(* IEC 61131-3 sources: daoli-st-library/DL_Process (part 2) *)

(* ---- FB_DL_ColumnDpCtrl.st ---- *)
(*==============================================================================
 * 组件名称 (Component)  : FB_DL_ColumnDpCtrl
 * 溯源说明 (Provenance): 道莅 clean-room 防御性实现（IEC 61131-3 纯净实现，闭源文档仅借语义，零代码行）
 * 所属子库 (Sublibrary) : DL_Process / ProcessControl
 * 当前版本 (Version)    : 1.0.0
 * 兼容性   (Platform)   : CODESYS 3.5 / TwinCAT 3 / 汇川 InoProShop / 施耐德
 *                         Machine Expert；纯 IEC 61131-3（第 3 版），仅用
 *                         Standard.library 的 TON / LIMIT / ABS / TIME_TO_DINT / DINT_TO_TIME
 * 组件分类 (Category)   : 功能块（FUNCTION_BLOCK）· 精馏塔压差控制
 * 功能一句话 (Summary)  : 以塔压差设定为基准增量式双向调节回流与再沸两路给定，
 *                         带死区、双侧抗饱和，压差越上限时按防冲塔策略强制分配。
 *
 * 本件存在的意义 (Why this unit exists)
 *   精馏塔的 ΔP 是「液泛前兆」的直接指示：ΔP 升高说明上升蒸汽被液相托住，
 *   继续加热会冲塔（产品全部跑废、可能超压）。库内 FB_DL_RatioController 管
 *   两路比值、FB_DL_SplitRangeControl 管单输出分程，都不解「ΔP 偏高时增回流
 *   减再沸、ΔP 偏低时反向」这条双向分配律，也没有防冲塔的强制优先级。
 *
 * 增量式调节与抗饱和 (Incremental law and anti-windup)
 *   两路输出都是**增量累加**的绝对给定（不是增量输出），每走一步：
 *     ΔP 偏高（> 设定 + 死区）→ 回流 +fStep、再沸 −fStep
 *     ΔP 偏低（< 设定 − 死区）→ 回流 −fStep、再沸 +fStep
 *   累加后钳到 fOutMin~fOutMax，且**到达限值即停止向该方向累加**——钳位后
 *   不再累加是本件的抗饱和手段，不做积分回算（塔的工艺时间常数以十分钟计，
 *   回算没有收益，只会让审计算不清）。
 *
 * 防冲塔优先级 (Anti-flooding priority)
 *   fDpMeas > fDpHighLimit 持续 tConfirm → bDpHigh：**再沸立即降到 fOutMin、
 *   回流抬到 fOutMax**，压差调节暂时让位。这条优先级高于增量调节，因为冲塔
 *   是不可逆的产品损失；退出须压差回落到 fDpHighLimit − fDpDeadband 以下
 *   （用已有死区引脚做回差，不新开参数），避免在限值上反复进出。
 *
 * 引脚补全声明 (Pin completion —— 规格正文要求但引脚表漏列)
 *   fStep : 单步调节量 [%]，规格正文明确要求「步长引脚 fStep（缺省 1.0 %）」；
 *   tStep : 步进节拍 [ms]，增量式调节必须有时基，否则步进率随任务周期漂移。
 *   tStep 采用 T#200MS 缺省（现场常规回路周期），两引脚均已按要求常量化默认值。
 *
 * 边界安全 (Boundary)
 *   ① fDpSp <= 0、fOutMin >= fOutMax、fDpHighLimit <= fDpSp、fStep <= 0、
 *      任一参数非有限 → 故障 030E、**双输出置 fOutMin**（切断热源侧再加量）；
 *   ② fDpMeas 非有限 → 故障 030F、**保持末次输出**（塔不能因坏值断热，
 *      与①方向相反，两条并列写死）；
 *   ③ 死区内 → 信息 01DC，不调节、输出保持；
 *   ④ bDpHigh 进入置 01DD，退出复用 01DC（R90 不加码，头注释写明复用理由）；
 *   ⑤ 失能 → eIdle、双输出置 fOutMin、bDpHigh 清零（逐项赋，R72）；
 *   ⑥ 两只 TON 无条件刷新（步进节拍 / 越限确认），各司其职不共用；
 *   ⑦ CASE 落 ELSE 置 0310 并回 eFault。
 *
 * 错误码    : 16#0005_01DC ΔP 在死区内不调节，或已退出防冲塔——信息级，正常调节
 *             16#0005_01DD ΔP 越上限，已按防冲塔策略强制分配——信息级，保护动作
 *             16#0005_030E 控制参数非法（设定/限值/步长/上下限关系）——故障级，双输出置下限
 *             16#0005_030F ΔP 输入非有限，保持末次输出——故障级，不得断热
 *             16#0005_0310 状态机落 ELSE 兜底（非法状态）——故障级，回 eFault
 * 码位总账  : 16#0005_01DC 用 / 16#0005_01DD 用 ｜ 16#0005_030E 用 / 16#0005_030F 用 / 16#0005_0310 用
 * 状态机    : E_DL_ColumnDpState（eIdle / eNormal / eDpHigh / eDpLow / eFault），CASE 含 ELSE 兜底，
 *             ELSE 置 16#0005_0310 并回 eFault；失能无条件回 eIdle
 * 采样约定  : 每任务周期调用一次；步进节拍由 tStep 给定，越限确认由 tConfirm 给定
 * 依赖说明  : 只做组合编排，不复制低层算法；无 DL_ 子库调用
 * 验收向量  : V1 ΔP 5.0、设定 5.0、死区 0.2 → 死区内不调节，eErr = 01DC，输出保持
 *             V2 ΔP 6.0（> 5.2）、步长 1.0、节拍 200 ms → 每步回流 +1、再沸 −1，
 *                累加到限值后停（抗饱和主向量）
 *             V3 V2 持续到回流 = fOutMax → bLimited = TRUE，不再向该方向累加
 *             V4 ΔP 8.5（> 上限 8.0）持续 2 s → bDpHigh = TRUE，回流 = fOutMax、
 *                再沸 = fOutMin，eErr = 01DD（防冲塔主向量）
 *             V5 V4 后 ΔP 回落到 7.9（< 8.0 − 0.2）→ 退出防冲塔，eErr = 01DC（回差主向量）
 *             V6 fDpSp = 0 → 030E，双输出 = fOutMin，bValid = FALSE
 *             V7 fDpMeas = NaN → 030F，双输出保持上一拍值（坏值不断热主向量）
 *             V8 bEnable 落 → eIdle，双输出 = fOutMin，bDpHigh = FALSE
 * 红线自检  : 全局变量声明零使用 / 外部变量访问零使用 / 物理地址零使用 ｜ 纯 IEC 61131-3 ｜ 无除法
 *             浮点只用大小与容差比较 ｜ 无循环 ｜ 全变量双语同行注释 ｜ ENUM + CASE
 *             含 ELSE ｜ 两只 TON 在主体前部无条件刷新 ｜ 阈值常量化，无魔法数
 * 修订历史  : 2026-11-16  v1.0.0  首版入库（R22 · 批 3 · 过程单元控制）
 *============================================================================*)

(*-----------------------------------------------------------------------------
 * 枚举: E_DL_ColumnDpState（归属本功能块，同文件发布，全库唯一定义）
 * 含义: 塔压差控制相位。0 起步长 10。
 *-----------------------------------------------------------------------------*)
TYPE E_DL_ColumnDpState :
(
    eIdle   := 0,      // 待机：未使能或参数非法 / Idle, disabled or illegal parameters
    eNormal := 10,     // 正常：ΔP 在死区外按增量调节 / Normal, incremental control outside the dead band
    eDpHigh := 20,     // 压差高：防冲塔强制分配 / High differential pressure, anti-flooding distribution
    eDpLow  := 30,     // 压差低：反向调节 / Low differential pressure, reverse correction
    eFault  := 99      // 故障：参数非法或输入非有限 / Fault, illegal parameter or non-finite input
);
END_TYPE

FUNCTION_BLOCK FB_DL_ColumnDpCtrl
VAR_INPUT
    fDpMeas      : REAL;                       // 塔压差实测 [kPa] / measured column differential pressure [kPa]
    fDpSp        : REAL := 5.0;                // 压差设定 [kPa]，须 > 0 / differential pressure setpoint [kPa], must be > 0
    fDpDeadband  : REAL := 0.2;                // 死区半宽 [kPa]，须 >= 0 / dead band half width [kPa], must be >= 0
    fOutMin      : REAL := 0.0;                // 输出下限 [%] / output floor [%]
    fOutMax      : REAL := 100.0;              // 输出上限 [%]，须 > fOutMin / output ceiling [%], must exceed the floor
    fDpHighLimit : REAL := 8.0;                // 防冲塔压差上限 [kPa]，须 > fDpSp / anti-flooding limit [kPa], must exceed the setpoint
    fStep        : REAL := 1.0;                // 单步调节量 [%]，须 > 0 / single step size [%], must be > 0
    tStep        : TIME := T#200MS;            // 步进节拍 [ms] / step cadence [ms]
    tConfirm     : TIME := T#2S;               // 越限确认时间 [ms] / limit confirm time [ms]
    bEnable      : BOOL;                       // 使能 / enable
END_VAR
VAR_OUTPUT
    fRefluxOut   : REAL;                       // 回流量给定 [%]，范围 fOutMin~fOutMax / reflux setpoint [%]
    fReboilOut   : REAL;                       // 再沸热源给定 [%]，范围 fOutMin~fOutMax / reboiler duty setpoint [%]
    bDpHigh      : BOOL;                       // 压差越上限（防冲塔生效） / differential pressure above the limit
    bLimited     : BOOL;                       // 输出已到限值（抗饱和生效） / an output sits at its limit
    eErr         : UDINT;                      // 错误码，0 表示无错 / error code, 0 means no error
    bError       : BOOL;                       // 故障级标志，仅故障级错误置位 / fault-class flag, set only on fault-level codes
    bValid       : BOOL;                       // 输出可用标志 / outputs usable flag
END_VAR
VAR
    fbStep       : TON;                        // 步进节拍计时，段 6 无条件刷新 [ms] / step cadence timer
    fbHigh       : TON;                        // 越限确认计时，段 6 无条件刷新 [ms] / limit confirm timer
    _eState      : E_DL_ColumnDpState := E_DL_ColumnDpState.eIdle; // 当前相位 / current phase
    _bInit       : BOOL := FALSE;              // 首扫标志，初值 FALSE 取非判定 / first-scan flag, tested negated
    _bParamBad   : BOOL;                       // 参数非法标志 / illegal parameter flag
    _bFiniteBad  : BOOL;                       // 输入非有限标志 / non-finite input flag
    _bIllegal    : BOOL;                       // 非法状态标志 / illegal state flag
    _bStepBreak  : BOOL;                       // 步进计时器断输入一拍 / step timer one-scan break
    _bHighBreak  : BOOL;                       // 越限计时器断输入一拍 / limit timer one-scan break
    _bStepPulse  : BOOL;                       // 本拍走一步 / one step this scan
    _bInDeadband : BOOL;                       // 本拍在死区内 / inside the dead band this scan
    _bHiAbove    : BOOL;                       // 本拍越上限（裸判据） / above the limit this scan
    _bHiExit     : BOOL;                       // 压差已回落到退出线以下 / below the exit line
    _tStepUse    : TIME := T#200MS;            // 生效步进节拍 [ms]，已钳位 / effective cadence, clamped
    _tConfUse    : TIME := T#2S;               // 生效确认时间 [ms]，已钳位 / effective confirm time, clamped
    _fReflux     : REAL;                       // 回流量累加保持量 [%] / held reflux setpoint [%]
    _fReboil     : REAL;                       // 再沸累加保持量 [%] / held reboiler setpoint [%]
    _fRefluxOut  : REAL;                       // 回流输出暂存 [%] / reflux outlet staging
    _fReboilOut  : REAL;                       // 再沸输出暂存 [%] / reboiler outlet staging
END_VAR
VAR CONSTANT
    DL_VAL_LIM     : REAL := 1.0E6;            // 有限性判定的绝对值上限 [无量纲] / finiteness ceiling
    DL_SP_MIN      : REAL := 0.0;              // 设定下限 [kPa]，须严格大于 / setpoint floor, strictly greater
    DL_BAND_MIN    : REAL := 0.0;              // 死区下限 [kPa] / dead band floor [kPa]
    DL_STEP_MIN    : REAL := 0.0;              // 步长下限 [%]，须严格大于 / step floor, strictly greater
    DL_EPS         : REAL := 1.0E-6;           // 浮点比较容差 [%] / float comparison tolerance [%]
    DL_CAD_MIN_MS  : DINT := 10;               // 步进节拍下限 [ms] / cadence floor [ms]
    DL_CAD_MAX_MS  : DINT := 60000;            // 步进节拍上限 [ms] / cadence ceiling [ms]
    DL_CONF_MAX_MS : DINT := 60000;            // 确认时间上限 [ms] / confirm ceiling [ms]
    DL_TIME_ZERO   : TIME := T#0MS;            // 时间零值基准 [ms] / time zero reference
END_VAR

(*------------------------------------------------------------------------------
 * 段 1｜每拍预置（输出与累加量在段 9 单点写入）
 *      Per-scan presets, the outputs and accumulators are written in segment nine
 *-----------------------------------------------------------------------------*)
eErr         := 16#0000_0000;                  // 错误码每拍重算 / error code recomputed every scan
bError       := FALSE;                         // 故障标志每拍重算 / fault flag recomputed every scan
bValid       := FALSE;                         // 可用标志每拍重算 / usable flag recomputed every scan
bDpHigh      := FALSE;                         // 越限标志每拍重算 / high flag recomputed
bLimited     := FALSE;                         // 抗饱和标志每拍重算 / limited flag recomputed
_bParamBad   := FALSE;                         // 参数非法标志预清零 / parameter flag pre-cleared
_bFiniteBad  := FALSE;                         // 非有限标志预清零 / non-finite flag pre-cleared
_bIllegal    := FALSE;                         // 非法状态标志预清零 / illegal state flag pre-cleared
_bStepPulse  := FALSE;                         // 步进脉冲预置 FALSE / step pulse preset FALSE
_bInDeadband := FALSE;                         // 死区标志预置 FALSE / dead band flag preset FALSE
_bHiAbove    := FALSE;                         // 越上限标志预置 FALSE / above-limit preset FALSE
_bHiExit     := FALSE;                         // 退出标志预置 FALSE / exit preset FALSE

(*------------------------------------------------------------------------------
 * 段 2｜首扫初始化（两路从输出下限起：塔未运行时回流与热源都在最小位）
 *      First-scan initialisation, both loops start at the output floor
 *-----------------------------------------------------------------------------*)
IF NOT _bInit THEN
    _eState     := E_DL_ColumnDpState.eIdle;   // 相位待机 / phase idle
    _fReflux    := 0.0;                        // 回流累加量 0 [%] / reflux accumulator zero
    _fReboil    := 0.0;                        // 再沸累加量 0 [%] / reboiler accumulator zero
    _bStepBreak := TRUE;                       // 步进节拍从零开始 / cadence timer starts from zero
    _bHighBreak := TRUE;                       // 越限确认从零开始 / confirm timer starts from zero
    _bInit      := TRUE;                       // 首扫只做一次 / the first scan runs once
END_IF

(*------------------------------------------------------------------------------
 * 段 3｜参数闸门（设定/上下限关系/越限值/步长，任一非法即故障级）
 *      Parameter gate, any illegal value or relation is a fault
 *-----------------------------------------------------------------------------*)
IF (fDpSp <> fDpSp) OR (ABS(fDpSp) > DL_VAL_LIM) OR (fDpSp <= DL_SP_MIN) THEN
    _bParamBad := TRUE;                        // 压差设定非法 / setpoint illegal
END_IF
IF (fOutMin <> fOutMin) OR (fOutMax <> fOutMax) OR (ABS(fOutMin) > DL_VAL_LIM)
   OR (ABS(fOutMax) > DL_VAL_LIM) THEN
    _bParamBad := TRUE;                        // 输出上下限非有限 / output limits non-finite
ELSIF fOutMin >= fOutMax THEN
    _bParamBad := TRUE;                        // 上下限关系非法 / illegal limit relation
END_IF
IF (fDpHighLimit <> fDpHighLimit) OR (ABS(fDpHighLimit) > DL_VAL_LIM)
   OR (fDpHighLimit <= fDpSp) THEN
    _bParamBad := TRUE;                        // 越限值必须严格大于设定 / the limit must exceed the setpoint
END_IF
IF (fStep <> fStep) OR (ABS(fStep) > DL_VAL_LIM) OR (fStep <= DL_STEP_MIN) THEN
    _bParamBad := TRUE;                        // 步长非法 / step illegal
END_IF
IF (fDpDeadband <> fDpDeadband) OR (fDpDeadband < DL_BAND_MIN) OR (ABS(fDpDeadband) > DL_VAL_LIM) THEN
    _bParamBad := TRUE;                        // 死区非法 / dead band illegal
END_IF

(*------------------------------------------------------------------------------
 * 段 4｜输入有限性（区间判据同时拦 NaN 与 ±Inf）
 *      Input finiteness, the interval test catches NaN and infinity
 *-----------------------------------------------------------------------------*)
IF (fDpMeas < -DL_VAL_LIM) OR (fDpMeas > DL_VAL_LIM) THEN
    _bFiniteBad := TRUE;                       // 压差非有限 / differential pressure non-finite
END_IF

(*------------------------------------------------------------------------------
 * 段 5｜判据计算（死区 / 越上限 / 退出线，全部在参数合法时才可信）
 *      Criteria evaluation, only meaningful with legal parameters
 *-----------------------------------------------------------------------------*)
IF (NOT _bFiniteBad) AND (NOT _bParamBad) THEN
    _bInDeadband := (ABS(fDpMeas - fDpSp) <= fDpDeadband); // 死区判据 [布尔] / dead band test
    _bHiAbove    := (fDpMeas > fDpHighLimit);              // 越上限裸判据 / raw above-limit test
    _bHiExit     := (fDpMeas < (fDpHighLimit - fDpDeadband)); // 退出线用已有死区做回差 / the exit line reuses the dead band
END_IF

(*------------------------------------------------------------------------------
 * 段 6｜两只计时器无条件刷新（R40：CASE 之外每拍必调，各司其职不共用）
 *      Both timers refreshed unconditionally, each with its own duty
 *-----------------------------------------------------------------------------*)
_tStepUse := tStep;                            // 步进节拍直取引脚 [ms] / cadence from the pin
IF TIME_TO_DINT(_tStepUse) < DL_CAD_MIN_MS THEN
    _tStepUse := DINT_TO_TIME(DL_CAD_MIN_MS);  // 下限钳位（无专用码位，R90 不新开码） / clamped to the floor
END_IF
IF TIME_TO_DINT(_tStepUse) > DL_CAD_MAX_MS THEN
    _tStepUse := DINT_TO_TIME(DL_CAD_MAX_MS);  // 上限钳位 / clamped to the ceiling
END_IF

_tConfUse := tConfirm;                         // 确认时间直取引脚 [ms] / confirm time from the pin
IF TIME_TO_DINT(_tConfUse) < 0 THEN
    _tConfUse := DL_TIME_ZERO;                 // 负时间兜底为 0 / fallback to zero
END_IF
IF TIME_TO_DINT(_tConfUse) > DL_CONF_MAX_MS THEN
    _tConfUse := DINT_TO_TIME(DL_CONF_MAX_MS); // 上限钳位 / clamped to the ceiling
END_IF

fbStep(IN := bEnable AND (NOT _bParamBad) AND (NOT _bFiniteBad)
             AND (NOT _bInDeadband) AND (NOT _bHiAbove) AND (NOT _bStepBreak),
       PT := _tStepUse);                       // 步进节拍计时
_bStepBreak := FALSE;                          // 断输入拍在调用后自清 / break self-cleared after the call
_bStepPulse := fbStep.Q;                       // 本拍走一步 / one step this scan

fbHigh(IN := bEnable AND (NOT _bParamBad) AND (NOT _bFiniteBad) AND _bHiAbove AND (NOT _bHighBreak),
       PT := _tConfUse);                       // 越限确认计时
_bHighBreak := FALSE;                          // 断输入拍在调用后自清 / break self-cleared after the call

(*------------------------------------------------------------------------------
 * 段 7｜相位机（只做迁移；调节量在段 8 演进）
 *      Phase machine, transitions only, the setpoints evolve in segment eight
 *-----------------------------------------------------------------------------*)
CASE _eState OF

    E_DL_ColumnDpState.eIdle:                  // 待机：参数合法且使能即进入
        IF _bParamBad OR _bFiniteBad THEN
            _eState := E_DL_ColumnDpState.eFault; // 原因未消失，转故障 / the cause persists
        ELSIF bEnable THEN
            IF fbHigh.Q THEN
                _eState := E_DL_ColumnDpState.eDpHigh; // 越限已确认，直接进防冲塔 / the limit is confirmed
                _bStepBreak := TRUE;           // 步进节拍重启 / the cadence restarts
            ELSIF (fDpSp - fDpMeas) > fDpDeadband THEN
                _eState := E_DL_ColumnDpState.eDpLow;  // 压差偏低，直接进低压相 / differential pressure low
            ELSE
                _eState := E_DL_ColumnDpState.eNormal; // 正常区间（含偏高与死区） / normal range
            END_IF
        END_IF

    E_DL_ColumnDpState.eNormal:                // 正常：越限或偏低都会迁移
        IF _bParamBad OR _bFiniteBad THEN
            _eState := E_DL_ColumnDpState.eFault; // 转故障 / go to fault
        ELSIF NOT bEnable THEN
            _eState := E_DL_ColumnDpState.eIdle;  // 失能回待机 / disabled, back to idle
        ELSIF fbHigh.Q THEN
            _eState := E_DL_ColumnDpState.eDpHigh; // 越限确认，进防冲塔 / confirmed, anti-flooding
            _bStepBreak := TRUE;               // 步进节拍重启 / the cadence restarts
        ELSIF (fDpSp - fDpMeas) > fDpDeadband THEN
            _eState := E_DL_ColumnDpState.eDpLow;  // 压差偏低 / differential pressure low
        END_IF

    E_DL_ColumnDpState.eDpLow:                 // 压差低：回升进死区即回正常
        IF _bParamBad OR _bFiniteBad THEN
            _eState := E_DL_ColumnDpState.eFault; // 转故障 / go to fault
        ELSIF NOT bEnable THEN
            _eState := E_DL_ColumnDpState.eIdle;  // 失能回待机 / disabled, back to idle
        ELSIF fbHigh.Q THEN
            _eState := E_DL_ColumnDpState.eDpHigh; // 越限确认，进防冲塔 / confirmed, anti-flooding
            _bStepBreak := TRUE;               // 步进节拍重启 / the cadence restarts
        ELSIF (fDpMeas - fDpSp) >= (-fDpDeadband) THEN
            _eState := E_DL_ColumnDpState.eNormal; // 已回到死区边界内 / back inside the dead band edge
        END_IF

    E_DL_ColumnDpState.eDpHigh:                // 防冲塔：压差回落到退出线以下才让位
        IF _bParamBad OR _bFiniteBad THEN
            _eState := E_DL_ColumnDpState.eFault; // 转故障 / go to fault
        ELSIF NOT bEnable THEN
            _eState := E_DL_ColumnDpState.eIdle;  // 失能回待机 / disabled, back to idle
        ELSIF _bHiExit THEN
            _eState := E_DL_ColumnDpState.eNormal; // 退出防冲塔（回差确认） / leave anti-flooding after hysteresis
            _bStepBreak := TRUE;               // 步进节拍重启，避免立即继续累加 / the cadence restarts
        END_IF

    E_DL_ColumnDpState.eFault:                 // 故障：参数与输入恢复即回待机
        IF bEnable AND (NOT _bParamBad) AND (NOT _bFiniteBad) THEN
            _eState := E_DL_ColumnDpState.eIdle; // 原因消失 / the cause is gone
            _bStepBreak := TRUE;               // 步进节拍重启 / the cadence restarts
        END_IF

    ELSE
        _bIllegal := TRUE;                     // 标记非法状态 / flag the illegal state
        _eState   := E_DL_ColumnDpState.eFault; // 回故障态 / back to the fault state
END_CASE

(*------------------------------------------------------------------------------
 * 段 8｜调节量演进（唯一累加点：防冲塔强制分配 > 步进增量）
 *      Setpoint evolution, the single accumulation point
 *-----------------------------------------------------------------------------*)
IF (_eState = E_DL_ColumnDpState.eDpHigh) AND (NOT _bFiniteBad) AND (NOT _bParamBad) THEN
    _fReflux := fOutMax;                       // 防冲塔：回流抬到上限 [%] / reflux forced to the ceiling
    _fReboil := fOutMin;                       // 防冲塔：再沸立即降到下限 [%] / reboiler forced to the floor
ELSIF _bStepPulse AND bEnable AND (NOT _bFiniteBad) AND (NOT _bParamBad)
      AND (_eState <> E_DL_ColumnDpState.eIdle) THEN
    IF (fDpMeas - fDpSp) > fDpDeadband THEN
        (* ΔP 偏高：增回流、减再沸，各自到达限值即停（抗饱和） *)
        (* High differential pressure, add reflux and cut reboiler, both stop at their limits *)
        IF _fReflux < (fOutMax - DL_EPS) THEN
            _fReflux := _fReflux + fStep;      // 回流增量 [%] / reflux increment
        END_IF
        IF _fReboil > (fOutMin + DL_EPS) THEN
            _fReboil := _fReboil - fStep;      // 再沸减量 [%] / reboiler decrement
        END_IF
    ELSIF (fDpSp - fDpMeas) > fDpDeadband THEN
        (* ΔP 偏低：减回流、增再沸，各自到达限值即停（抗饱和） *)
        (* Low differential pressure, cut reflux and add reboiler, both stop at their limits *)
        IF _fReflux > (fOutMin + DL_EPS) THEN
            _fReflux := _fReflux - fStep;      // 回流减量 [%] / reflux decrement
        END_IF
        IF _fReboil < (fOutMax - DL_EPS) THEN
            _fReboil := _fReboil + fStep;      // 再沸增量 [%] / reboiler increment
        END_IF
    END_IF
    _bStepBreak := TRUE;                       // 走一步后重启节拍，节拍严格等于 tStep / restart the cadence
END_IF

(* 限值钳位：参数变更或强制分配后一律落回 [fOutMin, fOutMax] *)
(* Clamped into the output range after any change *)
IF (NOT _bParamBad) THEN
    _fReflux := LIMIT(fOutMin, _fReflux, fOutMax); // 回流钳位 [%] / reflux clamped
    _fReboil := LIMIT(fOutMin, _fReboil, fOutMax); // 再沸钳位 [%] / reboiler clamped
END_IF

(*------------------------------------------------------------------------------
 * 段 9｜输出单点写入与码位优先级链
 *      Single write point of the outputs and the code priority chain
 *-----------------------------------------------------------------------------*)
IF _bParamBad THEN
    _fRefluxOut := fOutMin;                    // 参数非法：回流置下限（安全侧） [%] / reflux to the floor
    _fReboilOut := fOutMin;                    // 参数非法：再沸置下限（切断热源加量） [%] / reboiler to the floor
ELSIF NOT bEnable THEN
    _fRefluxOut := fOutMin;                    // 失能：回流置下限 [%] / reflux to the floor
    _fReboilOut := fOutMin;                    // 失能：再沸置下限 [%] / reboiler to the floor
ELSE
    _fRefluxOut := _fReflux;                   // 正常：回流给定 [%] / reflux setpoint
    _fReboilOut := _fReboil;                   // 正常：再沸给定 [%] / reboiler setpoint
END_IF

fRefluxOut := _fRefluxOut;                     // 回流出口 [%] / reflux outlet
fReboilOut := _fReboilOut;                     // 再沸出口 [%] / reboiler outlet
bDpHigh    := (_eState = E_DL_ColumnDpState.eDpHigh); // 越限标志出口 / high flag outlet
bLimited   := (_fRefluxOut >= (fOutMax - DL_EPS)) OR (_fRefluxOut <= (fOutMin + DL_EPS))
              OR (_fReboilOut >= (fOutMax - DL_EPS)) OR (_fReboilOut <= (fOutMin + DL_EPS)); // 任一输出到限值即置位

IF _bIllegal THEN
    eErr   := 16#0005_0310;                    // 故障级：状态机兜底 / fault: state machine fallback
    bError := TRUE;                            // 置故障标志 / raise the fault flag
ELSIF _bParamBad THEN
    eErr   := 16#0005_030E;                    // 故障级：控制参数非法 / fault: control parameters illegal
    bError := TRUE;                            // 置故障标志 / raise the fault flag
ELSIF _bFiniteBad THEN
    eErr   := 16#0005_030F;                    // 故障级：输入非有限，保持末次输出 / fault: non-finite input, outputs held
    bError := TRUE;                            // 置故障标志 / raise the fault flag
ELSIF bDpHigh THEN
    eErr   := 16#0005_01DD;                    // 信息级：越上限已按防冲塔策略分配 / informational: anti-flooding applied
ELSIF _bInDeadband THEN
    eErr   := 16#0005_01DC;                    // 信息级：死区内不调节（退出防冲塔亦复用本码） / informational: no correction
END_IF

IF bError THEN
    bValid := FALSE;                           // 故障级：输出不可用 / fault: outputs unusable
ELSIF NOT bEnable THEN
    bValid := FALSE;                           // 失能：输出不可用 / disabled: unusable
ELSE
    bValid := TRUE;                            // 输出可用 / outputs usable
END_IF

END_FUNCTION_BLOCK

(* ---- FB_DL_ConveyorMergePrioritySeq.st ---- *)
(*
  ============================================================
  组件名 : FB_DL_ConveyorMergePrioritySeq
  分类   : DL_Process
  功能   : 汇流合流优先权仲裁（主线优先、支线不饿死、抢占恢复、堵车计数告警、堵死与授权超时故障锁存）
  开源溯源 : internal-design（本轮无外部代码逐行引用）；参考语义 : 无外部参考
  复杂度 : C3
  版本   : 1.0.0
  ============================================================
*)

(*-----------------------------------------------------------------------------
 * 状态迁移表（ENUM 成员 → 出口；每成员均有可到达出口，零无界驻留相）：
 *   eIdle       → eGrantMain   : bReqMain（主线请求优先，含两路同时请求）
 *   eIdle       → eGrantBranch : 仅 bReqBranch 且无主线请求
 *   eIdle       ── 保持，直到任一请求（待机相以请求为唯一出口，属许可型驻留）
 *   eGrantMain  → eGrantBranch : bZoneMainClear 落沿（车辆已进入主线段，本次授权完成）且 bReqBranch
 *   eGrantMain  → eHoldBranch  : bZoneMainClear 落沿 且无支线请求（保持拦住支线）
 *   eGrantMain  → eJamWait     : bJamMain（主线堵车）
 *   eGrantMain  → eFault       : tonGrant.Q（码 2 单次授权超 tGrantMax）
 *   eGrantBranch→ eGrantMain   : bZoneBranchClear 落沿 且（抢占登记 或 主线再请求）
 *   eGrantBranch→ eIdle        : bZoneBranchClear 落沿 且无主线请求
 *   eGrantBranch→ eJamWait     : bJamBranch（支线堵车）
 *   eGrantBranch→ eFault       : tonGrant.Q（码 2 单次授权超 tGrantMax）
 *   eHoldBranch → eGrantMain   : bReqMain
 *   eHoldBranch → eGrantBranch : bReqBranch 且无主线请求
 *   eHoldBranch → eIdle        : 两路请求均已消失（进相前置条件消失，R98）
 *   eJamWait    → eIdle        : 对应堵车信号消失 ｜ rtJamReset.Q（bJamReset 上升沿）
 *   eJamWait    → eFault       : tonJamWait.Q（主线成因码 1 / 支线成因码 3）
 *   eFault      → eIdle        : bJamReset 上升沿（段 3 已清锁存，段 4 判锁存位迁相）
 *   ELSE（非法枚举值，非任何成员）→ eFault（码 5）
 *
 * 故障码表（nFaultCode，0 = 无故障；非首码均附「现有输出不可观测」反证句，R90）：
 *   1 主线堵死   : eJamWait 内主线堵车信号持续超 tJamTimeout（归因成员 _bJamFromMain = TRUE）。
 *   2 授权超时   : 反证——单次授权超 tGrantMax 时 eJamWait 未进入，堵车信号仍为假；
 *                  复用码 1 会把「光栅/清空信号失效」报成「物理堵料」，运维去拆包而非查光栅。
 *   3 支线堵死   : 反证——支线成因由 _bJamFromMain = FALSE 唯一标记，故障相动作全撤后
 *                  bGrantMainOut/bGrantBranchOut 同为 FALSE、eState 同为 eFault；若复用码 1，
 *                  运维将疏通主线而放过真正堵塞的支线（方向性误判，R146）。
 *   4 输入非法   : 反证——非有限速度或时间/计数参数越域时无任何请求沿、无授权动作，
 *                  与码 1/2/3 的时序签名互斥，必须独立成码以便组态错误可被前置拦截。
 *   5 非法状态   : 反证——非法枚举值为程序缺陷而非现场事件，合并入任一工艺码会让固件
 *                  错误被误排为设备故障，故独立成码。
 *
 * 依赖     : 仅 IEC 61131-3 标准库（TON / R_TRIG / F_TRIG / ABS），零厂商私有库
 * 分工声明 : 皮带驱动变频与速度环归驱动件；物理堵料检测（光电/限位）归现场检测件，
 *            本件只做「授权仲裁 + 堵车计数 + 安全撤权」，不做速度闭环也不做机械保护。
 * 归属     : E_DL_MergePrioState 归属本文件（全库唯一定义，R264；引用件只引用不重声明）。
 * 修订历史 : 2026-11-25  v1.0.0  首版（编码席 dlf-plc-coder，第二批 C3）
 *----------------------------------------------------------------------------*)

(*-----------------------------------------------------------------------------
 * 边界与红线自检：
 * ① 四个 TON 与三个沿实例（rtJamReset / ftMainClear / ftBranchClear）全部在 CASE 外无条件周期调用
 *    （R7）；时间类 IN 均含 NOT .Q 自复位项与 NOT 故障锁存项（R188 / FB50-1③），CASE 内只读 .Q。
 * ② 三个授权/保持出口在段 0 每拍预置 FALSE，CASE 内只置 TRUE —— eIdle 与 eFault 零残留。
 * ③ nJamCount 的写入点共三处且互不叠加：段 3 复位沿清零、eGrantMain/eGrantBranch 堵车事件入相 +1
 *    （一事件一次）、段 5 支线等待满窗 +1；不存在两处同拍 ±1 的双向计数（实战规则 1③）。
 * ④ 告警位 bJamAlarm 为纯派生式（计数超门槛 或 授权相内低速征兆），不独立锁存、无自引用赋值，
 *    计数被 bJamReset 清零后告警自动消失（R28 5.9 派生位纪律）。
 * ⑤ 堵车归因唯一：_bJamFromMain 在入相赋值点唯一，超时分支按该成员分列码 1 / 码 3（R190）。
 * ⑥ 复位沿作用域逐项声明（FB50-2②）：清堵车计数 / 清故障锁存与故障码 / 迁相回空闲，三项各写明。
 * ⑦ 低速征兆（|v| < 0.05）只参与告警计数，不单独触发故障（偏低类只降级，R146）。
 * ⑧ 零全局耦合：无 GVL / VAR_EXTERNAL / %I / %Q（R1 / R2）；无 FOR / WHILE / REPEAT（R271 N/A）。
 * ⑨ 相位写入点共两处且互斥：段 4 CASE、段 6 段尾迁移闸（无第三处旁路写相位）。
 *----------------------------------------------------------------------------*)

TYPE E_DL_MergePrioState :
(
    eIdle        := 0,                                              // 空闲：三路出口全撤，等请求 idle: all three outlets withdrawn, waiting for a request
    eGrantMain   := 1,                                              // 主线授权相：放行主线，支线请求挂起 main grant: main line released, branch requests parked
    eGrantBranch := 2,                                              // 支线授权相：放行支线，主线再请求时登记抢占 branch grant: branch released, a new main request registers preemption
    eHoldBranch  := 3,                                              // 支线保持拦截相：主线通过后拦住支线，等下一请求 hold branch: branch blocked after a main pass until the next request
    eJamWait     := 4,                                              // 堵车等待相：撤全部授权，等堵车信号消失或复位 jam wait: all grants withdrawn until the jam signal clears or a reset arrives
    eFault       := 5                                               // 故障锁存相：全部授权撤除，只由 bJamReset 沿迁出 fault: all grants withdrawn, left only by the bJamReset edge
);
END_TYPE

FUNCTION_BLOCK FB_DL_ConveyorMergePrioritySeq
VAR_INPUT
    bReqMain          : BOOL := FALSE;                              // 主线合流请求（电平）[bool] main line merge request level
    bReqBranch        : BOOL := FALSE;                              // 支线合流请求（电平）[bool] branch line merge request level
    bZoneMainClear    : BOOL := FALSE;                              // 主线段清空确认（TRUE = 段内无车）[bool] main segment clear confirmation, TRUE means empty
    bZoneBranchClear  : BOOL := FALSE;                              // 支线段清空确认（TRUE = 段内无车）[bool] branch segment clear confirmation, TRUE means empty
    bJamMain          : BOOL := FALSE;                              // 主线堵车检测（现场检测件给出）[bool] main line jam detection from the field device
    bJamBranch        : BOOL := FALSE;                              // 支线堵车检测（现场检测件给出）[bool] branch line jam detection from the field device
    rSpeedMain        : REAL := 0.0;                                // 主线实测线速度 [m/s] measured main line speed [m/s]
    rSpeedBranch      : REAL := 0.0;                                // 支线实测线速度 [m/s] measured branch line speed [m/s]
    tGrantMax         : TIME := T#30S;                              // 单次授权最长占用窗 [s] maximum single grant window [s]
    tJamTimeout       : TIME := T#60S;                              // 堵车持续判与支线等待计数窗 [s] jam persistence and branch wait counting window [s]
    nJamResetCountMax : INT := 3;                                   // 支线等待计数告警门槛，域 0..10000 [次] branch wait count alarm threshold, domain 0..10000
    bJamReset         : BOOL := FALSE;                              // 堵车复位（上升沿）：清计数与故障锁存 [bool] jam reset rising edge, clears the count and the fault latch
END_VAR
VAR_OUTPUT
    bGrantMainOut   : BOOL;                                         // 主线放行授权（段 0 预置，CASE 只置位）[bool] main line release grant
    bGrantBranchOut : BOOL;                                         // 支线放行授权（段 0 预置，CASE 只置位）[bool] branch line release grant
    bHoldBranchOut  : BOOL;                                         // 支线拦截保持（段 0 预置，CASE 只置位）[bool] branch line hold command
    eState          : E_DL_MergePrioState;                          // 相位出口（段 7 单点映射）[-] phase outlet mapped once in section 7
    nJamCount       : INT;                                          // 支线等待/堵车累计次数 [次] accumulated branch wait and jam event count
    bJamAlarm       : BOOL;                                         // 支线饥饿告警（计数派生，非故障）[bool] branch starvation alarm derived from the count, not a fault
    nFaultCode      : INT;                                          // 故障码 0 无 1 主线堵死 2 授权超时 3 支线堵死 4 输入非法 5 非法状态 [码] fault code
    bError          : BOOL;                                         // 故障锁存标志（取锁存位，R45 配对出口）[bool] fault latch flag used as the paired outlet
END_VAR
VAR
    _eState         : E_DL_MergePrioState := E_DL_MergePrioState.eIdle; // 内部相位（CASE 唯一比较目标）[-] internal phase compared by the CASE
    _bFaultLatch    : BOOL := FALSE;                                // 故障锁存位（仅 bJamReset 沿清除）[bool] fault latch, cleared only by the bJamReset edge
    _nFault         : INT := 0;                                     // 锁存故障码（故障期回放，不按当下输入重算）[码] latched fault code replayed in the fault phase
    _nJamCnt        : INT := 0;                                     // 内部支线等待与堵车计数 [次] internal branch wait and jam count
    _bCfgOk         : BOOL := FALSE;                                // 组态与入参域闸通过标志 [bool] configuration and input domain gate flag
    _bRunActive     : BOOL := FALSE;                                // 仲裁相关相标志（授权/保持/堵车等待）[bool] arbitration phase flag
    _bGrantMain     : BOOL := FALSE;                                // 内部主线授权状态 [bool] internal main grant state
    _bGrantBranch   : BOOL := FALSE;                                // 内部支线授权状态 [bool] internal branch grant state
    _bHoldBranch    : BOOL := FALSE;                                // 内部支线拦截状态 [bool] internal branch hold state
    _bPreemptPending : BOOL := FALSE;                               // 主线抢占登记（支线授权期间挂起）[bool] main preemption pending during a branch grant
    _bJamFromMain   : BOOL := TRUE;                                 // 堵车归因：TRUE 主线成因 / FALSE 支线成因（R190）[bool] jam attribution, TRUE for main and FALSE for branch
    _bSlowMain      : BOOL := FALSE;                                // 主线低速征兆（|v| < 门限）[bool] main line low speed symptom
    _bSlowBranch    : BOOL := FALSE;                                // 支线低速征兆（|v| < 门限）[bool] branch line low speed symptom
    rtJamReset      : R_TRIG;                                       // bJamReset 上升沿实例（段 2 无条件调用）[bool] jam reset rising edge instance
    ftMainClear     : F_TRIG;                                       // 主线段清空落沿实例（段 2 无条件调用）[bool] main segment clear falling edge instance
    ftBranchClear   : F_TRIG;                                       // 支线段清空落沿实例（段 2 无条件调用）[bool] branch segment clear falling edge instance
    tonGrant        : TON;                                          // 单次授权占用计时（段 2 无条件调用）[s] single grant occupancy timer
    tonJamWait      : TON;                                          // 堵车持续判计时（段 2 无条件调用）[s] jam persistence timer
    tonBranchWait   : TON;                                          // 支线等待满窗计数计时（段 2 无条件调用）[s] branch wait counting timer
END_VAR
VAR CONSTANT
    DL_MRG_ZERO      : REAL := 0.0;                                 // 浮点零基准 [m/s] float zero base
    DL_MRG_V_MIN     : REAL := 0.05;                                // 低速征兆门限 [m/s] low speed symptom threshold [m/s]
    DL_MRG_T_MIN     : TIME := T#100MS;                             // 时间参数下限 [s] lower bound of the time parameters
    DL_MRG_T_MAX     : TIME := T#2H;                                // 时间参数上限 [s] upper bound of the time parameters
    DL_MRG_CNT_MAX   : INT := 10000;                                // 计数门槛上限 [次] upper bound of the count threshold
    DL_MRG_CNT_ZERO  : INT := 0;                                    // 计数零基准 [次] count zero base
    DL_MRG_CNT_ONE   : INT := 1;                                    // 计数步长 [次] count step
END_VAR

(* —— 段 0：出口命令预置与派生量（CASE 内只置 TRUE，杜绝故障相残留） —— *)
_bGrantMain   := FALSE;                                             // 主线授权每拍先撤 [bool] main grant withdrawn first each scan
_bGrantBranch := FALSE;                                             // 支线授权每拍先撤 [bool] branch grant withdrawn first each scan
_bHoldBranch  := FALSE;                                             // 支线拦截每拍先撤 [bool] branch hold withdrawn first each scan
_bRunActive   := (_eState = E_DL_MergePrioState.eGrantMain) OR (_eState = E_DL_MergePrioState.eGrantBranch)
                 OR (_eState = E_DL_MergePrioState.eHoldBranch) OR (_eState = E_DL_MergePrioState.eJamWait); // 仲裁相标志（用状态量，R99）[bool] arbitration phase flag
_bSlowMain    := (ABS(rSpeedMain) < DL_MRG_V_MIN);                  // 主线低速征兆（非有限值此判恒假，由域闸兜住）[bool] main low speed symptom
_bSlowBranch  := (ABS(rSpeedBranch) < DL_MRG_V_MIN);                // 支线低速征兆（非有限值此判恒假，由域闸兜住）[bool] branch low speed symptom

(* —— 段 1：组态域闸（全部浮点入参与时间/计数参数枚举，非有限双判 R151 / R79） —— *)
_bCfgOk := TRUE;                                                    // 组态闸标志初值 [bool] configuration flag initial value
IF (rSpeedMain <> rSpeedMain) OR ((rSpeedMain - rSpeedMain) <> DL_MRG_ZERO)
   OR (rSpeedBranch <> rSpeedBranch) OR ((rSpeedBranch - rSpeedBranch) <> DL_MRG_ZERO) THEN
    _bCfgOk := FALSE;                                               // 非有限速度：拒收（NaN 自反 + Inf 差值自减）[bool] non finite speed rejected
END_IF
IF _bCfgOk THEN
    IF (tGrantMax < DL_MRG_T_MIN) OR (tGrantMax > DL_MRG_T_MAX) THEN
        _bCfgOk := FALSE;                                           // 授权窗越域 [bool] grant window out of domain
    ELSIF (tJamTimeout < DL_MRG_T_MIN) OR (tJamTimeout > DL_MRG_T_MAX) THEN
        _bCfgOk := FALSE;                                           // 堵车窗越域 [bool] jam window out of domain
    ELSIF (nJamResetCountMax < DL_MRG_CNT_ZERO) OR (nJamResetCountMax > DL_MRG_CNT_MAX) THEN
        _bCfgOk := FALSE;                                           // 告警门槛越域 [bool] alarm threshold out of domain
    END_IF
END_IF
IF (NOT _bCfgOk) AND (NOT _bFaultLatch) AND (bReqMain OR bReqBranch OR _bRunActive) THEN
    _nFault      := 4;                                              // 故障级：输入非法（非有限/越域）[码] fault: illegal input
    _bFaultLatch := TRUE;                                           // 置故障锁存 [bool] latch the fault
    bError       := TRUE;                                           // R45 配对：故障标志同拍置位 [bool] paired error flag
END_IF

(* —— 段 2：沿与定时器（CASE 外无条件周期调用，R7；IN 含 NOT .Q 自复位与 NOT 锁存，R188） —— *)
rtJamReset(CLK := bJamReset);                                       // 复位沿无条件刷新 [bool] reset edge refreshed unconditionally
ftMainClear(CLK := bZoneMainClear);                                 // 主线段清空落沿刷新 [bool] main clear falling edge refreshed
ftBranchClear(CLK := bZoneBranchClear);                             // 支线段清空落沿刷新 [bool] branch clear falling edge refreshed
tonGrant(IN := ((_eState = E_DL_MergePrioState.eGrantMain) OR (_eState = E_DL_MergePrioState.eGrantBranch))
              AND (NOT tonGrant.Q) AND (NOT _bFaultLatch),
         PT := tGrantMax);                                          // 单次授权占用计时 [s] single grant occupancy timer
tonJamWait(IN := (_eState = E_DL_MergePrioState.eJamWait) AND (NOT tonJamWait.Q) AND (NOT _bFaultLatch),
           PT := tJamTimeout);                                      // 堵车持续判计时 [s] jam persistence timer
tonBranchWait(IN := bReqBranch AND (NOT bReqMain)
                 AND ((_eState = E_DL_MergePrioState.eGrantMain) OR (_eState = E_DL_MergePrioState.eHoldBranch))
                 AND (NOT tonBranchWait.Q) AND (NOT _bFaultLatch),
              PT := tJamTimeout);                                   // 支线被拦等待满窗计数 [s] branch blocked wait counting timer

(* —— 段 3：复位沿优先消化（作用域逐项声明，FB50-2②；先消化沿再消化超时，R275） —— *)
IF rtJamReset.Q THEN
    _nJamCnt := DL_MRG_CNT_ZERO;                                    // 复位沿作用域①：清支线等待与堵车计数 [次] reset scope one, clear the wait count
    IF _bFaultLatch THEN
        _bFaultLatch := FALSE;                                      // 复位沿作用域②：清故障锁存 [bool] reset scope two, clear the fault latch
        _nFault      := 0;                                          // 复位沿作用域③：清故障码 [码] reset scope three, clear the fault code
    END_IF
END_IF

(* —— 段 4：主状态机（相位写入点之一；每成员独立标签，ELSE 只兜非法值，FB32-5） —— *)
CASE _eState OF
E_DL_MergePrioState.eIdle :                                         // 空闲相：三路出口已撤
    IF bReqMain THEN
        _bPreemptPending := FALSE;                                  // 新周期清抢占登记 [bool] clear the preemption flag for the new cycle
        _eState := E_DL_MergePrioState.eGrantMain;                  // 迁移：主线优先 [phase] main line has priority
    ELSIF bReqBranch THEN
        _bPreemptPending := FALSE;                                  // 新周期清抢占登记 [bool] clear the preemption flag for the new cycle
        _eState := E_DL_MergePrioState.eGrantBranch;                // 迁移：仅支线请求 [phase] branch request only
    END_IF

E_DL_MergePrioState.eGrantMain :                                    // 主线授权相
    _bGrantMain := TRUE;                                            // 放行主线 [bool] release the main line
    IF bJamMain THEN
        _bJamFromMain := TRUE;                                      // 归因：主线成因（唯一赋值点，R190）[bool] attribution to the main line
        _nJamCnt      := _nJamCnt + DL_MRG_CNT_ONE;                 // 一次堵车事件一次计数 [次] one count per jam event
        _eState       := E_DL_MergePrioState.eJamWait;              // 迁移：撤权进堵车等待 [phase] withdraw and wait for the jam to clear
    ELSIF ftMainClear.Q THEN
        IF bReqBranch THEN
            _eState := E_DL_MergePrioState.eGrantBranch;            // 迁移：主线段已进车，放行支线 [phase] main entry done, release the branch
        ELSE
            _eState := E_DL_MergePrioState.eHoldBranch;             // 迁移：无支线请求，保持拦住支线 [phase] no branch request, hold the branch
        END_IF
    END_IF

E_DL_MergePrioState.eGrantBranch :                                  // 支线授权相
    _bGrantBranch := TRUE;                                          // 放行支线 [bool] release the branch line
    IF bReqMain THEN
        _bPreemptPending := TRUE;                                   // 登记主线抢占（支线通过后立即恢复主线）[bool] register main preemption
    END_IF
    IF bJamBranch THEN
        _bJamFromMain := FALSE;                                     // 归因：支线成因（唯一赋值点，R190）[bool] attribution to the branch line
        _nJamCnt      := _nJamCnt + DL_MRG_CNT_ONE;                 // 一次堵车事件一次计数 [次] one count per jam event
        _eState       := E_DL_MergePrioState.eJamWait;              // 迁移：撤权进堵车等待 [phase] withdraw and wait for the jam to clear
    ELSIF ftBranchClear.Q THEN
        IF _bPreemptPending OR bReqMain THEN
            _bPreemptPending := FALSE;                              // 抢占已兑现，清登记 [bool] preemption honoured, clear the flag
            _eState := E_DL_MergePrioState.eGrantMain;              // 迁移：支线通过后恢复主线 [phase] branch passed, restore the main line
        ELSE
            _eState := E_DL_MergePrioState.eIdle;                   // 迁移：无主线请求回空闲重新仲裁 [phase] no main request, back to idle
        END_IF
    END_IF

E_DL_MergePrioState.eHoldBranch :                                   // 支线保持拦截相
    _bHoldBranch := TRUE;                                           // 保持拦住支线 [bool] hold the branch line
    IF bReqMain THEN
        _eState := E_DL_MergePrioState.eGrantMain;                  // 迁移（出口 1）：主线请求 [phase] main request arrives
    ELSIF bReqBranch THEN
        _eState := E_DL_MergePrioState.eGrantBranch;                // 迁移（出口 2）：仅支线请求，不再拦 [phase] branch only, stop holding
    ELSIF (NOT bReqMain) AND (NOT bReqBranch) THEN
        _eState := E_DL_MergePrioState.eIdle;                       // 迁移（出口 3）：进相前置条件消失 [phase] both requests gone, the hold precondition vanished
    END_IF

E_DL_MergePrioState.eJamWait :                                      // 堵车等待相：三路授权已撤
    IF rtJamReset.Q THEN
        _eState := E_DL_MergePrioState.eIdle;                       // 迁移（出口 1）：人工复位直接回空闲 [phase] manual reset back to idle
    ELSIF _bJamFromMain AND (NOT bJamMain) THEN
        _eState := E_DL_MergePrioState.eIdle;                       // 迁移（出口 2）：主线堵车信号消失 [phase] main jam signal gone
    ELSIF (NOT _bJamFromMain) AND (NOT bJamBranch) THEN
        _eState := E_DL_MergePrioState.eIdle;                       // 迁移（出口 3）：支线堵车信号消失 [phase] branch jam signal gone
    END_IF

E_DL_MergePrioState.eFault :                                        // 故障锁存相：三路授权已由段 6 全撤
    IF NOT _bFaultLatch THEN
        _eState := E_DL_MergePrioState.eIdle;                       // 复位沿已在段 3 清锁存，此处迁回空闲 [phase] the latch was cleared in section 3
    END_IF

ELSE                                                                // 非法枚举值兜底（R6 / FB32-5）
    IF NOT _bFaultLatch THEN
        _nFault      := 5;                                          // 故障级：非法状态枚举值 [码] fault: illegal state enum value
        _bFaultLatch := TRUE;                                       // 置故障锁存 [bool] latch the fault
        bError       := TRUE;                                       // R45 配对：故障标志同拍置位 [bool] paired error flag
    END_IF
    _eState := E_DL_MergePrioState.eFault;                          // 非法值一律落安全相 [phase] illegal value falls into the safe phase
END_CASE

(* —— 段 5：超时看门狗与支线等待计数（状态已迁出则该相看门狗不生效，R275） —— *)
IF tonGrant.Q AND (NOT _bFaultLatch)
   AND ((_eState = E_DL_MergePrioState.eGrantMain) OR (_eState = E_DL_MergePrioState.eGrantBranch)) THEN
    _nFault      := 2;                                              // 故障级：单次授权超时 [码] fault: single grant timeout
    _bFaultLatch := TRUE;                                           // 置故障锁存 [bool] latch the fault
    bError       := TRUE;                                           // R45 配对：故障标志同拍置位 [bool] paired error flag
END_IF
IF tonJamWait.Q AND (NOT _bFaultLatch) AND (_eState = E_DL_MergePrioState.eJamWait) THEN
    IF _bJamFromMain THEN
        _nFault := 1;                                               // 故障级：主线堵死 [码] fault: main line blocked
    ELSE
        _nFault := 3;                                               // 故障级：支线堵死 [码] fault: branch line blocked
    END_IF
    _bFaultLatch := TRUE;                                           // 置故障锁存 [bool] latch the fault
    bError       := TRUE;                                           // R45 配对：故障标志同拍置位 [bool] paired error flag
END_IF
IF tonBranchWait.Q AND (NOT _bFaultLatch) AND (NOT rtJamReset.Q) THEN
    _nJamCnt := _nJamCnt + DL_MRG_CNT_ONE;                          // 支线被拦满一个窗 → 累计一次（单点写入；复位沿同拍优先，R275）[次] one count per blocked window
END_IF

(* —— 段 6：段尾故障迁移闸 + 故障/空闲相授权全撤（FB50-1④） —— *)
IF _bFaultLatch AND (_eState <> E_DL_MergePrioState.eFault) THEN
    _eState := E_DL_MergePrioState.eFault;                          // 锁存即迁相（锁存与迁相分离，R21）[phase] a latch forces the fault phase
END_IF
IF (_eState = E_DL_MergePrioState.eFault) OR (_eState = E_DL_MergePrioState.eIdle)
   OR (_eState = E_DL_MergePrioState.eJamWait) THEN
    _bGrantMain   := FALSE;                                         // 安全侧：主线授权全撤 [bool] main grant withdrawn on the safe side
    _bGrantBranch := FALSE;                                         // 安全侧：支线授权全撤 [bool] branch grant withdrawn on the safe side
    _bHoldBranch  := FALSE;                                         // 安全侧：支线拦截全撤 [bool] branch hold withdrawn on the safe side
END_IF

(* —— 段 7：统一出口（相位映射 + 计数与告警派生 + 锁存码回放；告警为纯派生位，无独立锁存） —— *)
bGrantMainOut   := _bGrantMain;                                     // 主线授权出口 [bool] main grant outlet
bGrantBranchOut := _bGrantBranch;                                   // 支线授权出口 [bool] branch grant outlet
bHoldBranchOut  := _bHoldBranch;                                    // 支线拦截出口 [bool] branch hold outlet
eState          := _eState;                                         // 相位出口 [phase] phase outlet
nJamCount       := _nJamCnt;                                        // 计数出口 [次] count outlet
bJamAlarm       := ((_nJamCnt > nJamResetCountMax) AND (nJamResetCountMax >= DL_MRG_CNT_ZERO))
                   OR (((_eState = E_DL_MergePrioState.eGrantMain) AND _bSlowMain)
                       OR ((_eState = E_DL_MergePrioState.eGrantBranch) AND _bSlowBranch)); // 告警纯派生：计数超门槛 或 授权中低速征兆（R28 5.9）
nFaultCode      := _nFault;                                         // 故障码出口（锁存回放）[码] fault code outlet replayed from the latch
bError          := _bFaultLatch;                                    // 故障标志取锁存位 [bool] fault flag from the latch
END_FUNCTION_BLOCK

(* ---- FB_DL_DryerZoneProfileSeq.st ---- *)
(*
  ============================================================
  组件名 : FB_DL_DryerZoneProfileSeq
  分类   : DL_Process
  功能   : 多温区烘干升温曲线执行（预热 → 斜率限制升温 → 保温 → 冷却 → 完成），含超温退避、升温超时、区号越界、超温持续、人工停止、冷却超时六类保护
  开源溯源 : internal-design（本轮无外部代码逐行引用）；参考语义 : 无外部参考
  复杂度 : C4
  版本   : 1.0.0
  ============================================================
*)

(*-----------------------------------------------------------------------------
 * 状态迁移表（ENUM 成员 → 出口；每成员均有可到达出口，零无界驻留相）：
 *   eIdle     → ePreheat  : bStart 且 bStop = FALSE 且区号合法且组态闸通过
 *   eIdle     ── 保持，直到启动（待机相以启动命令为唯一出口，属许可型驻留）
 *   ePreheat  → eRampUp   : 全部有效区 aTempAct ≥ 目标×0.3 - 保温带 ｜ 超温退避（设定冻结）
 *   ePreheat  → eFault    : tonRamp.Q（码 1 升温超时）｜ rtStop.Q（码 4 人工停止）
 *   eRampUp   → eSoak     : 最冷区 aTempAct ≥ (目标 - 保温带) - 1E-6
 *   eRampUp   ── 超温退避时驻留本相（不退相，只撤加热并冻结 aTempSp，超温持续由码 3 兜底）
 *   eRampUp   → eFault    : tonRamp.Q（码 1）｜ tonOverTemp.Q（码 3）｜ rtStop.Q（码 4）
 *   eSoak     → eCoolDown : tonSoak.Q（保温时间到）
 *   eSoak     → eRampUp   : 超温退避（设定冻结后回升温相）
 *   eSoak     → eFault    : tonOverTemp.Q（码 3）｜ rtStop.Q（码 4）
 *   eCoolDown → eDone     : 最热区 aTempAct ≤ 目标×0.2 + 1E-6
 *   eCoolDown → eFault    : tonCool.Q（码 5 冷却超时）｜ rtStop.Q（码 4）
 *   eDone     → eIdle     : bStart 撤除 ｜ rtStop.Q（完成相撤令）
 *   eFault    → eIdle     : bStop 上升沿（清锁存、清全部设定与输出）
 *   ELSE（非法枚举值，非任何成员）→ eFault（码 7）
 *
 * 故障码表（nFaultCode，0 = 无故障；非首码均附「现有输出不可观测」反证句，R90）：
 *   1 升温超时   : tonRamp 覆盖 ePreheat + eRampUp（相序串行，进 ePreheat 时计时器自然复位）。
 *   2 区号越界   : 反证——区号越域时 aTempSp 全零、bHeaterEnable = FALSE，与码 1 的输出组合同形，
 *                  复用码 1 会把「组态写错温区数」报成「加热能力不足」，导致加功率的错误处置。
 *   3 超温持续   : 反证——bHeaterEnable 已由退避撤除、aTempSp 冻结，故障相动作全撤后与码 1 的
 *                  观测量一致；复用码 1 会掩盖「超温保护未及时动作」这一安全相关首因。
 *   4 人工停止   : 反证——操作员主动停机属安全审计事件，必须与设备异常分离，
 *                  否则无法在停机记录中区分人为与故障。
 *   5 冷却超时   : 反证——冷却相 bHeaterEnable = FALSE 且 bCoolFanEnable = TRUE，故障撤除后
 *                  与码 1 全同；复用码 1 会让运维去查加热回路而非冷却风机/水路。
 *   6 参数非法   : 反证——非法参数在启动瞬间即拦截，此时无加热、无爬升历史，
 *                  与任何超时码的时序签名互斥，必须独立成码。
 *   7 非法状态   : 反证——非法枚举值为程序缺陷而非工艺事件，合并入任一工艺码会让固件错误
 *                  被误排为现场故障，必须独立成码。
 *
 * 依赖     : 仅 IEC 61131-3 标准库（TON / R_TRIG / ABS / LIMIT），零厂商私有库
 * 代理节拍 : R95 三句声明——① 代理值为固定 100ms 爬升节拍（DL_DRY_DT），本件无采样周期引脚；
 *            ② 覆盖任务周期 ≤ 100ms 的常规配置；③ 任务周期 > 100ms 的区间由上层循环周期
 *            监视件负责，本件不做补偿（周期超限时爬升偏慢，属验收债项）。
 * 分工声明 : 各温区独立 PID 与加热功率分配归温区调节件；本件只输出区级温度设定曲线与
 *            加热/冷却使能，不做连续调节、不做风机电流保护。
 * 归属     : E_DL_DryerState 归属本文件（全库唯一定义，R264；引用件只引用不重声明）。
 * 修订历史 : 2026-11-25  v1.0.0  首版（编码席 dlf-plc-coder，第二批 C4）
 *----------------------------------------------------------------------------*)

(*-----------------------------------------------------------------------------
 * 边界与红线自检：
 * ① 五个 TON 与一个 R_TRIG 全部在 CASE 外无条件周期调用（R7）；时间类 IN 均含 NOT .Q 自复位项
 *    与 NOT 故障锁存项（R188 / FB50-1③），CASE 内只读 .Q。
 * ② aTempSp 是「保持槽」而非单拍量：段 7 统一出口按相映射，eIdle / eFault 相强制全零，
 *    且段 6 在故障/空闲相把内部曲线 _aSpRamp 一并清零 —— 上轮 MAJOR 型「故障后残留旧设定」已双重封堵。
 * ③ 超温退避（R191 显式声明）：段 6 撤加热但不迁相，aTempSp 冻结于当前值；超温持续超
 *    tOverTempLimit 才由 tonOverTemp 锁存码 3。段 5 判定序保证同拍时码 3 优先于码 1。
 * ④ 斜率限制：eRampUp 内 aTempSp 每 100ms 节拍只推进 rRampRate/60 × 0.1 K，并饱和到
 *    (目标 - 保温带)，不存在阶跃路径；未装区（下标 ≥ _nZoneClamp）恒写 0。
 * ⑤ 看门狗使能域（R145）：tonRamp / tonSoak / tonCool 的 IN 只取相驻留本身，不叠加业务条件补集。
 * ⑥ 三族循环（R271）：本件只用 FOR，逐对计数 FOR ↔ END_FOR 相等（交付前行数复核）。
 * ⑦ 组态域闸枚举全部浮点入参（含数组四个元素）：aTempAct[0..3] / rTempTarget / rRampRate /
 *    rSoakBand / rOverTempLimit，NaN 自反 + Inf 差值自减双判（R151 / R79）。
 * ⑧ 零全局耦合：无 GVL / VAR_EXTERNAL / %I / %Q（R1 / R2）。
 * ⑨ 相位写入点共两处且互斥：段 4 CASE、段 6 段尾迁移闸。
 *----------------------------------------------------------------------------*)

TYPE E_DL_DryerState :
(
    eIdle     := 0, // 空闲：加热与冷却全停，区级设定全零 idle: heater and fan off, all zone setpoints zero
    ePreheat  := 1, // 预热相：各区设定升至目标×0.3，加热使能 preheat: zone setpoints at 0.3 of the target, heater enabled
    eRampUp   := 2, // 升温相：按 rRampRate 斜率限制爬升 ramp up: climbing with the slope limited by rRampRate
    eSoak     := 3, // 保温相：设定保持目标温度等 tSoakTime soak: setpoints held at the target until tSoakTime elapses
    eCoolDown := 4, // 冷却相：关加热、开冷却风机，设定全零 cool down: heater off, cooling fan on, setpoints zero
    eFault    := 5, // 故障锁存相：加热与冷却全停，设定全零，只由 bStop 沿迁出 fault: all outputs off, left only by the bStop edge
    eDone     := 6  // 完成相：曲线结束，等撤令 done: profile finished, waiting for the start to be withdrawn
);
END_TYPE

FUNCTION_BLOCK FB_DL_DryerZoneProfileSeq
VAR_INPUT
    bStart          : BOOL := FALSE;                          // 启动/运行许可（电平）：撤除即回空闲 [bool] start and run permissive level
    bStop           : BOOL := FALSE;                          // 人工停止（上升沿）：运行中置码 4，故障相为复位沿 [bool] manual stop rising edge, code 4 while running and the reset edge in fault
    nZoneCount      : INT := 4;                               // 装机温区数，有效域 1..4 [区] installed zone count, valid domain 1..4
    aTempAct        : ARRAY[0..3] OF REAL;                    // 各区实测温度 [degC] measured temperature per zone [degC]
    rTempTarget     : REAL := 80.0;                           // 工艺目标温度，域 > 0 [degC] process target temperature, domain > 0 [degC]
    rRampRate       : REAL := 2.0;                             // 升温斜率，域 > 0 [K/min] ramp rate, domain > 0 [K/min]
    rSoakBand       : REAL := 2.0;                            // 保温带（升温转保温的余量），域 ≥ 0 [K] soak band used by the ramp to soak transition [K]
    tSoakTime       : TIME := T#30M;                          // 保温时长 [s] soak duration [s]
    rOverTempLimit  : REAL := 100.0;                          // 超温保护门限，域 > rTempTarget [degC] over temperature limit, domain above the target [degC]
    tRampTimeout    : TIME := T#60M;                          // 预热+升温总超时窗，亦作冷却超时窗 [s] preheat and ramp timeout, also used by the cooling phase
    tOverTempLimit  : TIME := T#10S;                          // 超温持续判故障窗 [s] over temperature persistence window before the fault [s]
END_VAR
VAR_OUTPUT
    aTempSp          : ARRAY[0..3] OF REAL;                   // 各区温度设定曲线（段 7 统一映射，空闲/故障相强制全零）[degC] zone setpoint profile forced to zero in idle and fault
    eState           : E_DL_DryerState;                       // 相位出口（段 7 单点映射）[-] phase outlet mapped once in section 7
    bHeaterEnable    : BOOL;                                  // 加热总使能（超温退避与故障/空闲相强制 FALSE）[bool] heater master enable forced off on retreat and in idle/fault
    bCoolFanEnable   : BOOL;                                  // 冷却风机使能（仅冷却相）[bool] cooling fan enable, cooling phase only
    bOverTempAlarm   : BOOL;                                  // 超温告警（本体超温 或 超温故障锁存派生）[bool] over temperature alarm derived from the condition or the latched code
    bDone            : BOOL;                                  // 曲线完成（由相位派生，非单拍脉冲）[bool] profile done derived from the phase as a level
    nFaultCode       : INT;                                   // 故障码 0 无 1 升温超时 2 区号越界 3 超温持续 4 人工停止 5 冷却超时 6 参数非法 7 非法状态 [码] fault code
    rRampProgressPct : REAL;                                  // 最冷区温度相对目标的完成度 0..100 [%] coldest zone temperature versus target in percent [%]
    bError           : BOOL;                                  // 故障锁存标志（取锁存位，R45 配对出口）[bool] fault latch flag used as the paired outlet
END_VAR
VAR
    _eState       : E_DL_DryerState := E_DL_DryerState.eIdle;  // 内部相位（CASE 唯一比较目标）[-] internal phase compared by the CASE
    _bFaultLatch  : BOOL := FALSE;                             // 故障锁存位（仅 bStop 沿清除）[bool] fault latch, cleared only by the bStop edge
    _nFault       : INT := 0;                                  // 锁存故障码（故障期回放，不按当下输入重算）[码] latched fault code replayed in the fault phase
    _bCfgOk       : BOOL := FALSE;                             // 组态与入参域闸通过标志 [bool] configuration and input domain gate flag
    _bRunActive   : BOOL := FALSE;                             // 曲线执行相标志（预热到冷却）[bool] profile running phase flag from preheat to cool down
    _bHeater      : BOOL := FALSE;                             // 内部加热使能状态 [bool] internal heater enable state
    _bCoolFan     : BOOL := FALSE;                             // 内部冷却风机状态 [bool] internal cooling fan state
    _bOverTemp    : BOOL := FALSE;                             // 任一有效区超温标志 [bool] any active zone over the limit
    _aSpRamp      : ARRAY[0..3] OF REAL;                       // 内部区级设定保持槽（保持槽，非单拍量）[degC] internal zone setpoint holding slots
    _nZoneClamp   : INT := 1;                                  // 区数钳位值 1..4 [区] clamped zone count
    _nIdx         : INT := 0;                                  // 区遍历下标（FOR 专用）[区] zone loop index
    _rMinAct      : REAL := 0.0;                               // 有效区实测温度最小值（最冷区）[degC] minimum measured temperature of the active zones [degC]
    _rMaxAct      : REAL := 0.0;                               // 有效区实测温度最大值（最热区）[degC] maximum measured temperature of the active zones [degC]
    _rPreheatSp   : REAL := 0.0;                               // 预热设定 = 目标 × 0.3 [degC] preheat setpoint at 0.3 of the target [degC]
    _rCoolSp      : REAL := 0.0;                               // 冷却终点 = 目标 × 0.2 [degC] cooling end point at 0.2 of the target [degC]
    _rRampCeil    : REAL := 0.0;                               // 升温上限 = 目标 - 保温带 [degC] ramp ceiling at the target minus the soak band [degC]
    _rStep        : REAL := 0.0;                               // 单个节拍的爬升增量 [K] ramp increment of one tick [K]
    _rDtStep      : REAL := 0.0;                               // 本拍节拍秒数（非节拍拍为 0）[s] tick seconds of this scan, zero on non tick scans [s]
    _rProg        : REAL := 0.0;                               // 完成度中间量 [%] progress intermediate value [%]
    rtStop        : R_TRIG;                                    // bStop 上升沿实例（段 2 无条件调用）[bool] stop rising edge instance
    tonDtTick     : TON;                                       // 爬升节拍发生器（段 2 无条件调用，IN := NOT .Q 自复位）[s] ramp tick generator with self reset
    tonRamp       : TON;                                       // 预热+升温总超时计时（段 2 无条件调用）[s] preheat and ramp timeout
    tonSoak       : TON;                                       // 保温时长计时（段 2 无条件调用）[s] soak duration timer
    tonCool       : TON;                                       // 冷却超时计时（段 2 无条件调用）[s] cooling timeout timer
    tonOverTemp   : TON;                                       // 超温持续计时（段 2 无条件调用）[s] over temperature persistence timer
END_VAR
VAR CONSTANT
    DL_DRY_ZERO          : REAL := 0.0;      // 浮点零基准 [degC] float zero base
    DL_DRY_ONE           : REAL := 1.0;      // 浮点一基准 [-] float one base
    DL_DRY_HUNDRED       : REAL := 100.0;    // 百分比满量程 [%] percent full scale
    DL_DRY_SIXTY         : REAL := 60.0;     // 每分钟秒数（K/min → K/s 换算）[s] seconds per minute for the K/min conversion
    DL_DRY_EPS           : REAL := 1.0E-6;   // 温度比较容差 [K] temperature comparison tolerance
    DL_DRY_PREHEAT_RATIO : REAL := 0.3;      // 预热比例（目标×0.3）[-] preheat ratio of the target
    DL_DRY_COOL_RATIO    : REAL := 0.2;      // 冷却终点比例（目标×0.2）[-] cooling end ratio of the target
    DL_DRY_DT_SEC        : REAL := 0.1;      // 爬升节拍秒数 [s] ramp tick length in seconds
    DL_DRY_DT            : TIME := T#100MS;  // 爬升节拍周期 [s] ramp tick period
    DL_DRY_IDX_MIN       : INT := 1;         // 区下标起点（下标 0 由初值行处理）[区] zone index start whose index zero is handled by the initialisation line
    DL_DRY_ZONE_MAX      : INT := 3;         // 区下标上限（定长数组上界）[区] zone index upper bound of the fixed array
    DL_DRY_ZONE_CNT_MAX  : INT := 4;         // 温区数上限（定长数组元素个数）[区] zone count upper bound of the fixed array
    DL_DRY_T_MIN         : TIME := T#100MS;  // 时间参数下限 [s] lower bound of the time parameters
    DL_DRY_T_MAX         : TIME := T#8H;     // 时间参数上限 [s] upper bound of the time parameters
END_VAR

(* —— 段 0：安全侧出口预置、区数钳位、温度极值与超温判据（CASE 只置 TRUE / 只推进曲线） —— *)
_bHeater   := FALSE;                                                // 加热使能每拍先撤（CASE 内只置 TRUE）[bool] heater withdrawn first each scan
_bCoolFan  := FALSE;                                                // 冷却风机每拍先撤（CASE 内只置 TRUE）[bool] cooling fan withdrawn first each scan
_rProg     := DL_DRY_ZERO;                                          // 完成度中间量每拍清零 [%] progress intermediate cleared each scan
_nZoneClamp := LIMIT(DL_DRY_IDX_MIN, nZoneCount, DL_DRY_ZONE_CNT_MAX); // 区数钳位 1..4（数组下标安全）[区] clamp the zone count
_rPreheatSp := rTempTarget * DL_DRY_PREHEAT_RATIO;                  // 预热设定 = 目标 × 0.3 [degC] preheat setpoint
_rCoolSp    := rTempTarget * DL_DRY_COOL_RATIO;                     // 冷却终点 = 目标 × 0.2 [degC] cooling end point
_rRampCeil  := rTempTarget - rSoakBand;                             // 升温上限 = 目标 - 保温带 [degC] ramp ceiling
IF _rRampCeil < DL_DRY_ZERO THEN
    _rRampCeil := DL_DRY_ZERO;                                      // 上限负值钳零（防负爬升目标）[degC] clamp a negative ceiling to zero
END_IF
_rMinAct   := aTempAct[0];                                          // 最冷区初值取下标 0 [degC] coldest zone seeded with index zero
_rMaxAct   := aTempAct[0];                                          // 最热区初值取下标 0 [degC] hottest zone seeded with index zero
_bOverTemp := (aTempAct[0] > rOverTempLimit);                       // 下标 0 的超温判据 [bool] over temperature check of index zero
FOR _nIdx := DL_DRY_IDX_MIN TO DL_DRY_ZONE_MAX DO
    IF _nIdx < _nZoneClamp THEN
        IF aTempAct[_nIdx] < _rMinAct THEN
            _rMinAct := aTempAct[_nIdx];                            // 刷新最冷区 [degC] refresh the coldest zone
        END_IF
        IF aTempAct[_nIdx] > _rMaxAct THEN
            _rMaxAct := aTempAct[_nIdx];                            // 刷新最热区 [degC] refresh the hottest zone
        END_IF
        IF aTempAct[_nIdx] > rOverTempLimit THEN
            _bOverTemp := TRUE;                                     // 任一有效区超温 [bool] any active zone over the limit
        END_IF
    END_IF
END_FOR
_bRunActive := (_eState = E_DL_DryerState.ePreheat) OR (_eState = E_DL_DryerState.eRampUp)
               OR (_eState = E_DL_DryerState.eSoak) OR (_eState = E_DL_DryerState.eCoolDown); // 曲线执行相标志（用状态量，R99）[bool] profile running flag

(* —— 段 1：组态域闸（浮点入参含数组四元素全枚举；区号越界独立成员判定，R151 / R79） —— *)
_bCfgOk := TRUE;                                                    // 组态闸标志初值 [bool] configuration flag initial value
IF (aTempAct[0] <> aTempAct[0]) OR ((aTempAct[0] - aTempAct[0]) <> DL_DRY_ZERO)
   OR (aTempAct[1] <> aTempAct[1]) OR ((aTempAct[1] - aTempAct[1]) <> DL_DRY_ZERO)
   OR (aTempAct[2] <> aTempAct[2]) OR ((aTempAct[2] - aTempAct[2]) <> DL_DRY_ZERO)
   OR (aTempAct[3] <> aTempAct[3]) OR ((aTempAct[3] - aTempAct[3]) <> DL_DRY_ZERO)
   OR (rTempTarget <> rTempTarget) OR ((rTempTarget - rTempTarget) <> DL_DRY_ZERO)
   OR (rRampRate <> rRampRate) OR ((rRampRate - rRampRate) <> DL_DRY_ZERO)
   OR (rSoakBand <> rSoakBand) OR ((rSoakBand - rSoakBand) <> DL_DRY_ZERO)
   OR (rOverTempLimit <> rOverTempLimit) OR ((rOverTempLimit - rOverTempLimit) <> DL_DRY_ZERO) THEN
    _bCfgOk := FALSE;                                               // 非有限入参：拒收（NaN 自反 + Inf 差值自减）[bool] non finite input rejected
END_IF
IF (bStart OR _bRunActive) AND (NOT _bFaultLatch) THEN
    IF (nZoneCount < DL_DRY_IDX_MIN) OR (nZoneCount > DL_DRY_ZONE_CNT_MAX) THEN
        _nFault      := 2;                                          // 故障级：区号越界（独立成因，R190）[码] fault: zone count out of domain
        _bFaultLatch := TRUE;                                       // 置故障锁存 [bool] latch the fault
        bError       := TRUE;                                       // R45 配对：故障标志同拍置位 [bool] paired error flag
    ELSE
        IF (NOT _bCfgOk) THEN
            _nFault      := 6;                                      // 故障级：参数非法（非有限/越域）[码] fault: illegal parameter
            _bFaultLatch := TRUE;                                   // 置故障锁存 [bool] latch the fault
            bError       := TRUE;                                   // R45 配对：故障标志同拍置位 [bool] paired error flag
        ELSIF (rTempTarget <= DL_DRY_ZERO) OR (rRampRate <= DL_DRY_ZERO) THEN
            _nFault      := 6;                                      // 故障级：目标或斜率非正 [码] fault: non positive target or ramp rate
            _bFaultLatch := TRUE;                                   // 置故障锁存 [bool] latch the fault
            bError       := TRUE;                                   // R45 配对：故障标志同拍置位 [bool] paired error flag
        ELSIF (rSoakBand < DL_DRY_ZERO) OR (rSoakBand >= rTempTarget) THEN
            _nFault      := 6;                                      // 故障级：保温带越域 [码] fault: soak band out of domain
            _bFaultLatch := TRUE;                                   // 置故障锁存 [bool] latch the fault
            bError       := TRUE;                                   // R45 配对：故障标志同拍置位 [bool] paired error flag
        ELSIF rOverTempLimit <= rTempTarget THEN
            _nFault      := 6;                                      // 故障级：超温门限不高于目标（必然误报）[码] fault: over temperature limit not above the target
            _bFaultLatch := TRUE;                                   // 置故障锁存 [bool] latch the fault
            bError       := TRUE;                                   // R45 配对：故障标志同拍置位 [bool] paired error flag
        ELSIF (tSoakTime < DL_DRY_T_MIN) OR (tSoakTime > DL_DRY_T_MAX) THEN
            _nFault      := 6;                                      // 故障级：保温时长越域 [码] fault: soak time out of domain
            _bFaultLatch := TRUE;                                   // 置故障锁存 [bool] latch the fault
            bError       := TRUE;                                   // R45 配对：故障标志同拍置位 [bool] paired error flag
        ELSIF (tRampTimeout < DL_DRY_T_MIN) OR (tRampTimeout > DL_DRY_T_MAX) THEN
            _nFault      := 6;                                      // 故障级：升温超时越域 [码] fault: ramp timeout out of domain
            _bFaultLatch := TRUE;                                   // 置故障锁存 [bool] latch the fault
            bError       := TRUE;                                   // R45 配对：故障标志同拍置位 [bool] paired error flag
        ELSIF (tOverTempLimit < DL_DRY_T_MIN) OR (tOverTempLimit > DL_DRY_T_MAX) THEN
            _nFault      := 6;                                      // 故障级：超温持续窗越域 [码] fault: over temperature window out of domain
            _bFaultLatch := TRUE;                                   // 置故障锁存 [bool] latch the fault
            bError       := TRUE;                                   // R45 配对：故障标志同拍置位 [bool] paired error flag
        END_IF
    END_IF
END_IF

(* —— 段 2：沿、定时器与节拍推进（CASE 外无条件周期调用，R7；IN 含 NOT .Q 自复位，R188） —— *)
rtStop(CLK := bStop);                                               // bStop 边沿无条件刷新 [bool] stop edge refreshed unconditionally
tonDtTick(IN := NOT tonDtTick.Q, PT := DL_DRY_DT);                  // 爬升节拍发生器（自复位周期窗）[s] self resetting ramp tick
_rDtStep := DL_DRY_ZERO;                                            // 非节拍拍增量秒数置零 [s] zero tick seconds on non tick scans
IF tonDtTick.Q THEN
    _rDtStep := DL_DRY_DT_SEC;                                      // 节拍拍推进 0.1s [s] advance 0.1 s on a tick scan
END_IF
tonRamp(IN := ((_eState = E_DL_DryerState.ePreheat) OR (_eState = E_DL_DryerState.eRampUp))
              AND (NOT tonRamp.Q) AND (NOT _bFaultLatch),
        PT := tRampTimeout);                                        // 预热+升温总超时（只看相驻留，R145）[s] preheat and ramp timeout on dwell only
tonSoak(IN := (_eState = E_DL_DryerState.eSoak) AND (NOT tonSoak.Q) AND (NOT _bFaultLatch),
        PT := tSoakTime);                                           // 保温时长 [s] soak duration
tonCool(IN := (_eState = E_DL_DryerState.eCoolDown) AND (NOT tonCool.Q) AND (NOT _bFaultLatch),
        PT := tRampTimeout);                                        // 冷却超时（同一时间引脚，两窗相序串行不重叠）[s] cooling timeout sharing the same pin
tonOverTemp(IN := _bOverTemp AND (_eState <> E_DL_DryerState.eIdle) AND (NOT tonOverTemp.Q)
                AND (NOT _bFaultLatch),
            PT := tOverTempLimit);                                  // 超温持续计时 [s] over temperature persistence

(* —— 段 3：人工停止优先消化（置锁存不写相位，迁相由段 6，R21 / R275） —— *)
IF rtStop.Q AND _bRunActive AND (NOT _bFaultLatch) THEN
    _nFault      := 4;                                              // 故障级：人工停止 [码] fault: manual stop
    _bFaultLatch := TRUE;                                           // 置故障锁存 [bool] latch the fault
    bError       := TRUE;                                           // R45 配对：故障标志同拍置位 [bool] paired error flag
END_IF

(* —— 段 4：主状态机（相位写入点之一；每成员独立标签，ELSE 只兜非法值，FB32-5） —— *)
CASE _eState OF
E_DL_DryerState.eIdle :                                             // 空闲相：设定与输出全零
    FOR _nIdx := 0 TO DL_DRY_ZONE_MAX DO
        _aSpRamp[_nIdx] := DL_DRY_ZERO;                             // 空闲相曲线保持槽清零（防空闲残留）[degC] clear the holding slots while idle
    END_FOR
    IF bStart AND (NOT bStop) AND _bCfgOk AND (NOT _bFaultLatch) THEN
        _eState := E_DL_DryerState.ePreheat;                        // 迁移：进入预热相 [phase] move to preheat
    END_IF

E_DL_DryerState.ePreheat :                                          // 预热相：各区设定 = 目标×0.3
    _bHeater := TRUE;                                               // 加热使能 [bool] heater enabled
    FOR _nIdx := 0 TO DL_DRY_ZONE_MAX DO
        IF _nIdx < _nZoneClamp THEN
            _aSpRamp[_nIdx] := _rPreheatSp;                         // 有效区写预热设定 [degC] active zone preheat setpoint
        ELSE
            _aSpRamp[_nIdx] := DL_DRY_ZERO;                         // 未装区恒零 [degC] uninstalled zone forced to zero
        END_IF
    END_FOR
    IF _bOverTemp THEN
        _eState := E_DL_DryerState.eRampUp;                         // 迁移：超温退避回升温相（设定冻结，加热由段 6 撤）[phase] retreat to ramp up
    ELSIF _rMinAct >= (_rPreheatSp - rSoakBand) THEN
        _eState := E_DL_DryerState.eRampUp;                         // 迁移：全部有效区达预热温度 [phase] preheat temperature reached
    END_IF

E_DL_DryerState.eRampUp :                                           // 升温相：斜率限制爬升（核心相）
    _bHeater := TRUE;                                               // 加热使能 [bool] heater enabled
    IF NOT _bOverTemp THEN
        _rStep := (rRampRate * _rDtStep) / DL_DRY_SIXTY;            // K/min × 节拍秒 / 60 → 单节拍增量 [K] per tick increment
        FOR _nIdx := 0 TO DL_DRY_ZONE_MAX DO
            IF _nIdx < _nZoneClamp THEN
                IF (_aSpRamp[_nIdx] + _rStep) < _rRampCeil THEN
                    _aSpRamp[_nIdx] := _aSpRamp[_nIdx] + _rStep;    // 斜率限制推进 [degC] slope limited advance
                ELSE
                    _aSpRamp[_nIdx] := _rRampCeil;                  // 饱和到升温上限（无阶跃超调）[degC] saturate at the ramp ceiling
                END_IF
            ELSE
                _aSpRamp[_nIdx] := DL_DRY_ZERO;                     // 未装区恒零 [degC] uninstalled zone forced to zero
            END_IF
        END_FOR
    END_IF
    IF (NOT _bOverTemp) AND (_rMinAct >= (_rRampCeil - DL_DRY_EPS)) THEN
        _eState := E_DL_DryerState.eSoak;                           // 迁移：最冷区到目标-保温带且未超温（防超温期抖动迁移）[phase] coldest zone reached the ceiling
    END_IF

E_DL_DryerState.eSoak :                                             // 保温相：设定保持目标温度
    _bHeater := TRUE;                                               // 加热使能 [bool] heater enabled
    FOR _nIdx := 0 TO DL_DRY_ZONE_MAX DO
        IF _nIdx < _nZoneClamp THEN
            _aSpRamp[_nIdx] := rTempTarget;                         // 有效区保温设定 = 目标 [degC] active zone soak setpoint
        ELSE
            _aSpRamp[_nIdx] := DL_DRY_ZERO;                         // 未装区恒零 [degC] uninstalled zone forced to zero
        END_IF
    END_FOR
    IF _bOverTemp THEN
        _eState := E_DL_DryerState.eRampUp;                         // 迁移：超温退避回升温相（设定冻结）[phase] retreat to ramp up
    ELSIF tonSoak.Q THEN
        _eState := E_DL_DryerState.eCoolDown;                       // 迁移：保温时间到 [phase] soak time elapsed
    END_IF

E_DL_DryerState.eCoolDown :                                         // 冷却相：关加热、开冷却风机
    _bCoolFan := TRUE;                                              // 冷却风机使能 [bool] cooling fan enabled
    FOR _nIdx := 0 TO DL_DRY_ZONE_MAX DO
        _aSpRamp[_nIdx] := DL_DRY_ZERO;                             // 冷却无加热需求，设定全零 [degC] no heating demand while cooling
    END_FOR
    IF _rMaxAct <= (_rCoolSp + DL_DRY_EPS) THEN
        _eState := E_DL_DryerState.eDone;                           // 迁移：最热区降到目标×0.2 [phase] hottest zone cooled down
    END_IF

E_DL_DryerState.eDone :                                             // 完成相：bDone 由相位派生
    FOR _nIdx := 0 TO DL_DRY_ZONE_MAX DO
        _aSpRamp[_nIdx] := DL_DRY_ZERO;                             // 完成相设定全零 [degC] setpoints zero after completion
    END_FOR
    IF (NOT bStart) OR rtStop.Q THEN
        _eState := E_DL_DryerState.eIdle;                           // 迁移：撤令或按停止回空闲 [phase] withdrawn start or a stop press returns to idle
    END_IF

E_DL_DryerState.eFault :                                            // 故障锁存相：输出与设定已由段 6 全撤
    FOR _nIdx := 0 TO DL_DRY_ZONE_MAX DO
        _aSpRamp[_nIdx] := DL_DRY_ZERO;                             // 故障相曲线保持槽清零 [degC] clear the holding slots in fault
    END_FOR
    IF rtStop.Q THEN
        _bFaultLatch := FALSE;                                      // 复位出口：清故障锁存 [bool] clear the fault latch
        _nFault      := 0;                                          // 复位出口：清故障码 [码] clear the fault code
        _eState      := E_DL_DryerState.eIdle;                      // 复位出口：迁回空闲（次拍 bStop 仍为 TRUE 不会误启动）[phase] back to idle
    END_IF

ELSE                                                                // 非法枚举值兜底（R6 / FB32-5）
    IF NOT _bFaultLatch THEN
        _nFault      := 7;                                          // 故障级：非法状态枚举值 [码] fault: illegal state enum value
        _bFaultLatch := TRUE;                                       // 置故障锁存 [bool] latch the fault
        bError       := TRUE;                                       // R45 配对：故障标志同拍置位 [bool] paired error flag
    END_IF
    _eState := E_DL_DryerState.eFault;                              // 非法值一律落安全相 [phase] illegal value falls into the safe phase
END_CASE

(* —— 段 5：超时看门狗锁存（判定序：超温持续优先于升温超时，同拍时码 3 优先，R190 归因唯一） —— *)
IF tonOverTemp.Q AND (NOT _bFaultLatch) AND (_eState <> E_DL_DryerState.eIdle) THEN
    _nFault      := 3;                                              // 故障级：超温持续 [码] fault: sustained over temperature
    _bFaultLatch := TRUE;                                           // 置故障锁存 [bool] latch the fault
    bError       := TRUE;                                           // R45 配对：故障标志同拍置位 [bool] paired error flag
END_IF
IF tonRamp.Q AND (NOT _bFaultLatch)
   AND ((_eState = E_DL_DryerState.ePreheat) OR (_eState = E_DL_DryerState.eRampUp)) THEN
    _nFault      := 1;                                              // 故障级：升温超时 [码] fault: ramp timeout
    _bFaultLatch := TRUE;                                           // 置故障锁存 [bool] latch the fault
    bError       := TRUE;                                           // R45 配对：故障标志同拍置位 [bool] paired error flag
END_IF
IF tonCool.Q AND (NOT _bFaultLatch) AND (_eState = E_DL_DryerState.eCoolDown) THEN
    _nFault      := 5;                                              // 故障级：冷却超时 [码] fault: cooling timeout
    _bFaultLatch := TRUE;                                           // 置故障锁存 [bool] latch the fault
    bError       := TRUE;                                           // R45 配对：故障标志同拍置位 [bool] paired error flag
END_IF
IF (NOT _bCfgOk) AND (NOT _bFaultLatch) AND _bRunActive THEN
    _nFault      := 6;                                              // 故障级：运行中出现非有限测量 [码] fault: non finite measurement during the run
    _bFaultLatch := TRUE;                                           // 置故障锁存 [bool] latch the fault
    bError       := TRUE;                                           // R45 配对：故障标志同拍置位 [bool] paired error flag
END_IF

(* —— 段 6：超温退避动作 + 段尾故障迁移闸 + 故障/空闲相动作与曲线全撤（FB50-1④） —— *)
IF _bOverTemp AND (_eState <> E_DL_DryerState.eFault) THEN
    _bHeater := FALSE;                                              // 超温退避：撤加热但不迁相（设定冻结，R191 显式声明）[bool] retreat: heater off without a phase change
END_IF
IF _bFaultLatch AND (_eState <> E_DL_DryerState.eFault) THEN
    _eState := E_DL_DryerState.eFault;                              // 锁存即迁相（锁存与迁相分离，R21）[phase] a latch forces the fault phase
END_IF
IF ((NOT bStart) AND _bRunActive AND (NOT _bFaultLatch)) OR (_eState = E_DL_DryerState.eFault) THEN
    (* 撤令语义（R191 二选一，本件选「降级为安全值 + 回空闲，不置故障码」）：加热与风机全停、曲线清零 *)
    IF (NOT bStart) AND (NOT _bFaultLatch)
       AND ((_eState = E_DL_DryerState.ePreheat) OR (_eState = E_DL_DryerState.eRampUp)
            OR (_eState = E_DL_DryerState.eSoak) OR (_eState = E_DL_DryerState.eCoolDown)) THEN
        _eState := E_DL_DryerState.eIdle;                           // 撤令即安全停机回空闲（用当拍相位判，不误吞 eDone）[phase] withdrawn start stops safely into idle
    END_IF
    _bHeater  := FALSE;                                             // 安全侧：加热全停 [bool] heater off on the safe side
    _bCoolFan := FALSE;                                             // 安全侧：冷却风机全停 [bool] cooling fan off on the safe side
    FOR _nIdx := 0 TO DL_DRY_ZONE_MAX DO
        _aSpRamp[_nIdx] := DL_DRY_ZERO;                             // 安全侧：曲线保持槽全零 [degC] clear all holding slots
    END_FOR
END_IF
IF _eState = E_DL_DryerState.eIdle THEN
    _bHeater  := FALSE;                                             // 空闲相：加热全停 [bool] heater off while idle
    _bCoolFan := FALSE;                                             // 空闲相：风机全停 [bool] cooling fan off while idle
    FOR _nIdx := 0 TO DL_DRY_ZONE_MAX DO
        _aSpRamp[_nIdx] := DL_DRY_ZERO;                             // 空闲相：曲线保持槽全零 [degC] clear all holding slots while idle
    END_FOR
END_IF

(* —— 段 7：统一出口（曲线映射 + 使能映射 + 完成度 + 锁存码回放；单点写入） —— *)
FOR _nIdx := 0 TO DL_DRY_ZONE_MAX DO
    IF (_eState = E_DL_DryerState.eIdle) OR (_eState = E_DL_DryerState.eFault)
       OR (_eState = E_DL_DryerState.eDone) THEN
        aTempSp[_nIdx] := DL_DRY_ZERO;                              // 空闲/故障/完成相：设定强制全零（MAJOR 型残留的双保险）[degC] setpoints forced to zero
    ELSE
        aTempSp[_nIdx] := _aSpRamp[_nIdx];                          // 运行相：映射内部曲线保持槽 [degC] map the internal holding slots
    END_IF
END_FOR
IF (rTempTarget > DL_DRY_EPS) AND _bCfgOk THEN
    _rProg := LIMIT(DL_DRY_ZERO, (_rMinAct * DL_DRY_HUNDRED) / rTempTarget, DL_DRY_HUNDRED); // 最冷区完成度（除子已双检，R4）[%] coldest zone progress
END_IF
bHeaterEnable    := _bHeater AND (_eState <> E_DL_DryerState.eIdle) AND (_eState <> E_DL_DryerState.eFault); // 加热使能出口（空闲/故障相强制 FALSE）[bool] heater enable outlet
bCoolFanEnable   := _bCoolFan AND (_eState <> E_DL_DryerState.eIdle) AND (_eState <> E_DL_DryerState.eFault); // 冷却风机出口（空闲/故障相强制 FALSE）[bool] cooling fan outlet
bOverTempAlarm   := _bOverTemp OR (_nFault = 3);                    // 超温告警：本体超温 或 超温故障锁存派生 [bool] over temperature alarm
eState           := _eState;                                        // 相位出口 [phase] phase outlet
bDone            := (_eState = E_DL_DryerState.eDone);               // 完成位由相位派生（非单拍脉冲）[bool] done derived from the phase
nFaultCode       := _nFault;                                        // 故障码出口（锁存回放）[码] fault code outlet replayed from the latch
rRampProgressPct := _rProg;                                         // 完成度出口 [%] progress outlet
bError           := _bFaultLatch;                                   // 故障标志取锁存位 [bool] fault flag from the latch
END_FUNCTION_BLOCK

(* ---- FB_DL_ElectrolyteFifoTrace.st ---- *)
(*==============================================================================
 * 组件名称 (Component)  : FB_DL_ElectrolyteFifoTrace
 * 所属子库 (Sublibrary) : DL_Process
 * 当前版本 (Version)    : 1.0.0
 * 兼容性   (Platform)   : CODESYS 3.5+ / TwinCAT 3 / 汇川 InoProShop / 施耐德 Machine Expert
 *                         仅依赖 Standard.library（R_TRIG / LEN / MUX 类标准函数），零厂商私有库
 * 功能描述 (Function)   : 注液批次 FIFO 追溯队列。
 *                         每支电芯注液完成时把"批次号 + 条码 + 注液量"三元组压入定长环形队列，
 *                         下游追溯/贴标工位按"先入先出"逐条取走，形成可回溯的注液履历链。
 *                         三条固化纪律：
 *                           ① **防重复入队**：压入前线性扫描在队记录，条码已存在即拒入（同一条码
 *                              在队列内只许出现一次，防重扫/重触发造成履历重复计数）；
 *                           ② **队满拒入**：计数达深度上限即拒入并锁存 bQueueFull，
 *                              直到出队使计数下降（或复位沿）才解除；
 *                           ③ **空队不宣称**：出队沿命中空队时 bOutValid=FALSE、不输出旧记录，
 *                              并按信息级置 eEmptyPop（不进锁存，R41 空队语义）。
 *                         验收向量：
 *                           ① 深度 32；压入 32 条后第 33 条 → 拒入 + bQueueFull 锁存
 *                           ② 同一 sBarcode 连续压入两次 → 第二次拒入 + eDupBarcode（不锁存）
 *                           ③ 空队出队 → bOutValid=FALSE + eEmptyPop（不锁存、不搬旧值）
 *                           ④ 满队后出队 1 条 → bQueueFull 解除，可再压入 1 条
 * 接口     (Interface)  : 入 bPush 入队沿、sBatchNo 批次号、sBarcode 电芯条码、fVolumeMl 注液量、
 *                         bPop 出队沿、bClear 清队沿、bReset 复位沿；
 *                         出 iQueueCnt 在队条数、sOutBatch / sOutBarcode / fOutVolumeMl 出队记录、
 *                         bOutValid 出队脉冲（单拍）、bQueueFull 队满锁存、bRejected 当拍拒入、
 *                         eState 相、eCause 成因、bError 故障标志。
 * 边界     (Boundary)   : ① **属主边界（写死）：本件只做"队列与履历记账"，不驱动注液泵/称重/
 *                         贴标机**，也不判注液量是否合格（属注液量判据件）；
 *                         ② **条码空串拒入**：LEN(sBarcode) = 0 → 拒入 + eBarcodeEmpty（信息级）；
 *                         ③ **深度闸**：环形指针一律以深度常量取模前先钳（下标恒在 1..32），
 *                         扫描循环带 _uGuard 计数器（上界 = 深度 + 2），循环必然收敛；
 *                         ④ **锁存解除式**：bQueueFull 的解除有两条——① 出队使计数 < 深度
 *                         （每拍重算，非沿）；② bReset 上升沿。两式自证可满足：出队沿与复位沿
 *                         均为外部引脚，不受任何锁存量门控，恒可达（R152/R234）；
 *                         ⑤ 组态/内部一致性故障（指针越界）→ 清队重建 + 锁存 ePtrCorrupt；
 *                         ⑥ 零全局耦合、零物理地址。
 * 分工声明 (Scope)      : 本件只管"注液履历队列"。不接管：注液量趋势判据
 *                         （属 FB_DL_ElectrolyteDosingTrend）、批次配方下发（属配方件）、
 *                         队列持久化落盘（属 MES 通讯件）。
 * 来源标签 (Source Tag) : ROADMAP 空勾真缺口 P1（注液批次追溯，自研 clean-room）
 * 码表     (Codes)      : 本件不占用任何全局数字码位（零码位范式 R297）；诊断由 BOOL + ENUM 出口承担。
 * 红线自检 (Redline)    : R1 ✓ 零 GVL/VAR_EXTERNAL ｜ R2 ✓ 零 %I/%Q/%M ｜ R3 ✓ 纯 IEC 61131-3
 *                         R4 ✓ 下标钳位 + 循环计数器 + 空串闸 + 满闸 ｜ R5 ✓ 声明逐行同行双语注释
 *                         R6 ✓ ENUM+CASE 含 ELSE 兜底 ｜ R7 ✓ R_TRIG 段 0 无条件刷新（本件无 TON）
 * 修订历史 (Revision)   : 2026-11-19  v1.0.0  R47 首版（批次 2 · 序号 6）
 *==============================================================================*)

TYPE ST_DL_EftRecord :
STRUCT
    sBatchNo  : STRING[31] := '';   // 注液批次号（≤31 字符） [-] / Electrolyte batch number, up to 31 chars
    sBarcode  : STRING[63] := '';   // 电芯条码（≤63 字符，队列内唯一） [-] / Cell barcode, unique inside the queue
    fVolumeMl : LREAL := 0.0;       // 本次注液量 [ml] / Injected volume of this shot [ml]
END_STRUCT
END_TYPE

TYPE E_DL_EftState :
(
    eIdle  := 0,    // 待机相（队列可用） / Idle, queue serviceable
    eFault := 90    // 故障相（指针损坏，等复位） / Fault, pointer corruption, awaiting reset
);
END_TYPE

TYPE E_DL_EftCause :
(
    eNone        := 0,   // 无异常 / No anomaly
    eDupBarcode  := 1,   // 条码重复（拒入，信息级） / Duplicate barcode, info level
    eBarcodeEmpty:= 2,   // 条码空串（拒入，信息级） / Empty barcode, info level
    eEmptyPop    := 3,   // 空队出队（不宣称，信息级） / Pop on empty queue, info level
    eQueueFull   := 4,   // 队满拒入（锁存） / Queue full, latched
    ePtrCorrupt  := 5,   // 环形指针损坏（故障级） / Ring pointer corruption, fault level
    ePhaseBad    := 6    // 非法相位兜底 / Illegal phase fallback
);
END_TYPE

FUNCTION_BLOCK FB_DL_ElectrolyteFifoTrace
VAR_INPUT
    bPush     : BOOL := FALSE;      // 入队沿 [-] / Enqueue edge
    sBatchNo  : STRING[31] := '';   // 待入队批次号 [-] / Batch number to enqueue
    sBarcode  : STRING[63] := '';   // 待入队电芯条码（队列内须唯一） [-] / Barcode to enqueue, unique inside the queue
    fVolumeMl : LREAL := 0.0;       // 待入队注液量 [ml] / Volume to enqueue [ml]
    bPop      : BOOL := FALSE;      // 出队沿 [-] / Dequeue edge
    bClear    : BOOL := FALSE;      // 清队沿（运维用，非故障路径） [-] / Clear edge, maintenance only
    bReset    : BOOL := FALSE;      // 故障复位沿 [-] / Fault reset edge
END_VAR
VAR_OUTPUT
    iQueueCnt    : INT := 0;                        // 在队条数 [条] / Records currently queued
    sOutBatch    : STRING[31] := '';                // 出队记录批次号 [-] / Dequeued batch number
    sOutBarcode  : STRING[63] := '';                // 出队记录条码 [-] / Dequeued barcode
    fOutVolumeMl : LREAL := 0.0;                    // 出队记录注液量 [ml] / Dequeued volume [ml]
    bOutValid    : BOOL := FALSE;                   // 出队脉冲（单拍，空队不宣称） [-] / Dequeue pulse, empty queue not claimed
    bQueueFull   : BOOL := FALSE;                   // 队满锁存 [-] / Queue full, latched
    bRejected    : BOOL := FALSE;                   // 当拍发生拒入 [-] / A push was rejected this scan
    bFullRelease : BOOL := FALSE;                   // 队满解除脉冲（单拍，诊断用） [-] / Full-release pulse, diagnostic
    eState       : E_DL_EftState := E_DL_EftState.eIdle;   // 相出口 [-] / Phase outlet
    eCause       : E_DL_EftCause := E_DL_EftCause.eNone;   // 成因出口（R190 归因唯一） [-] / Cause outlet
    bError       : BOOL := FALSE;                   // 故障标志（仅指针损坏级） [-] / Error flag, pointer corruption only
END_VAR
VAR
    _eState   : E_DL_EftState := E_DL_EftState.eIdle;      // 内部相（CASE 唯一写入目标） / Internal phase
    _eCause   : E_DL_EftCause := E_DL_EftCause.eNone;      // 成因锁存量 / Latched cause
    _bFault   : BOOL := FALSE;                             // 故障锁存位 / Latched fault bit
    _bFull    : BOOL := FALSE;                             // 队满锁存位（与 bQueueFull 同源） / Latched full bit
    _iHead    : INT := 1;                                  // 出队头指针（1..32） / Dequeue head pointer
    _iTail    : INT := 1;                                  // 入队尾指针（1..32） / Enqueue tail pointer
    _iCnt     : INT := 0;                                  // 在队条数 / Queued record count
    _bOutValid: BOOL := FALSE;                             // 出队脉冲内部位（单拍） / Internal dequeue pulse
    _bRejected: BOOL := FALSE;                             // 当拍拒入内部位（单拍） / Internal reject flag
    _bFullRel : BOOL := FALSE;                             // 队满解除内部位（单拍） / Internal full-release flag
    _bDup     : BOOL := FALSE;                             // 重复条码扫描结论 / Duplicate-scan result
    _uScan    : UINT := 0;                                 // 查重扫描计数器（防死循环） / Duplicate-scan guard counter
    _iScanIdx : INT := 0;                                  // 查重扫描下标（1..32） / Duplicate-scan index
    _bPushed  : BOOL := FALSE;                             // 本拍入队成功标志 / Push-succeeded flag of this scan
    rtPush    : R_TRIG;                                    // 入队沿实例，段 0 无条件调用 / Enqueue edge instance
    rtPop     : R_TRIG;                                    // 出队沿实例，段 0 无条件调用 / Dequeue edge instance
    rtClear   : R_TRIG;                                    // 清队沿实例，段 0 无条件调用 / Clear edge instance
    rtReset   : R_TRIG;                                    // 复位沿实例，段 0 无条件调用 / Reset edge instance
    aRec      : ARRAY[1..32] OF ST_DL_EftRecord;           // 记录环（深度字面量上界，R104） / Record ring, literal depth
END_VAR
VAR CONSTANT
    DL_EFT_DEPTH : INT := 32;           // 队列深度（与数组字面量上界同源，改动须同步） [条] / Queue depth
    DL_EFT_GUARD : UINT := 34;          // 查重循环守护上限（深度 + 2） [次] / Duplicate-scan guard limit
END_VAR

(* —— 段 0：四枚沿实例无条件周期刷新（R228A） —— *)
rtPush(CLK := bPush);                                       // 入队沿 / Enqueue edge
rtPop(CLK := bPop);                                         // 出队沿 / Dequeue edge
rtClear(CLK := bClear);                                     // 清队沿 / Clear edge
rtReset(CLK := bReset);                                     // 复位沿 / Reset edge

(* —— 段 1：单拍量预清零（锁存量 _eCause/_bFault/_bFull 不入清单，R107） —— *)
_bOutValid := FALSE;                                        // 出队脉冲预清 / Dequeue pulse preset
_bRejected := FALSE;                                        // 拒入标志预清 / Reject flag preset
_bFullRel  := FALSE;                                        // 满解除脉冲预清 / Full-release pulse preset
bError     := FALSE;                                        // 故障标志预清（R45 配对） / Error preset

(* —— 段 2：环形指针自检（越界即判损坏：清队重建 + 锁存） —— *)
IF (_iHead < 1) OR (_iHead > DL_EFT_DEPTH) OR (_iTail < 1) OR (_iTail > DL_EFT_DEPTH)
   OR (_iCnt < 0) OR (_iCnt > DL_EFT_DEPTH) THEN
    _iHead  := 1;                                           // 头指针重建 / Head rebuilt
    _iTail  := 1;                                           // 尾指针重建 / Tail rebuilt
    _iCnt   := 0;                                           // 计数清零 / Count cleared
    _eCause := E_DL_EftCause.ePtrCorrupt;                   // 归因：指针损坏 / Cause: pointer corruption
    _bFault := TRUE;                                        // 锁存 / Latch
    _eState := E_DL_EftState.eFault;                        // 入故障相 / Enter fault phase
END_IF

(* —— 段 3：迁出链（bReset 上升沿；bClear 为该沿之外的运维清队路径） —— *)
IF rtReset.Q THEN
    _bFault := FALSE;                                       // 清故障锁存 / Clear fault latch
    _bFull  := FALSE;                                       // 清队满锁存 / Clear full latch
    _eCause := E_DL_EftCause.eNone;                         // 清成因 / Clear cause
    _eState := E_DL_EftState.eIdle;                         // 回待机相 / Back to idle
END_IF
IF rtClear.Q THEN
    _iHead := 1;                                            // 头指针回 1 / Head back to 1
    _iTail := 1;                                            // 尾指针回 1 / Tail back to 1
    _iCnt  := 0;                                            // 计数清零 / Count cleared
    _bFull := FALSE;                                        // 清队满锁存 / Clear full latch
END_IF

(* —— 段 4：相迁移（故障相由段 3 迁出；本件无多相业务，故两相 CASE） —— *)
CASE _eState OF

E_DL_EftState.eIdle:
    ;                                                       // 待机相：队列服务在段 5/6 执行 / Service happens in stages 5 and 6

E_DL_EftState.eFault:
    ;                                                       // 故障相：仅等复位 / Wait for the reset edge only

ELSE
    _eCause := E_DL_EftCause.ePhaseBad;                     // 归因：非法相位 / Cause: illegal phase
    _bFault := TRUE;                                        // 锁存 / Latch
    _eState := E_DL_EftState.eFault;                        // 强拉故障相 / Force fault phase

END_CASE

(* —— 段 5：出队（FIFO 头指针推进；空队不宣称、不搬旧值） —— *)
IF (rtPop.Q) AND (_eState = E_DL_EftState.eIdle) THEN
    IF _iCnt > 0 THEN
        sOutBatch    := aRec[_iHead].sBatchNo;               // 取头记录批次号 / Take the head batch number
        sOutBarcode  := aRec[_iHead].sBarcode;               // 取头记录条码 / Take the head barcode
        fOutVolumeMl := aRec[_iHead].fVolumeMl;              // 取头记录注液量 / Take the head volume
        aRec[_iHead].sBatchNo  := '';                        // 清空已出队槽位批次号 / Clear the dequeued slot batch
        aRec[_iHead].sBarcode  := '';                        // 清空已出队槽位条码 / Clear the dequeued slot barcode
        aRec[_iHead].fVolumeMl := 0.0;                       // 清空已出队槽位注液量 / Clear the dequeued slot volume
        _bOutValid := TRUE;                                  // 出队脉冲 / Dequeue pulse
        _iCnt := _iCnt - 1;                                  // 计数递减 / Count decrement
        _iHead := _iHead + 1;                                // 头指针推进 / Head advance
        IF _iHead > DL_EFT_DEPTH THEN
            _iHead := 1;                                     // 环形回卷 / Ring wrap
        END_IF
        IF _bFull THEN
            _bFull := FALSE;                                 // 出队腾出空间：解除队满 / Space freed, clear the full latch
            _bFullRel := TRUE;                               // 满解除脉冲 / Full-release pulse
        END_IF
    ELSE
        _eCause := E_DL_EftCause.eEmptyPop;                  // 归因：空队出队（信息级，不锁存） / Cause: empty pop, info level
    END_IF
END_IF

(* —— 段 6：入队（先查重、再判满；拒入不改变队列内容） —— *)
IF (rtPush.Q) AND (_eState = E_DL_EftState.eIdle) THEN
    IF LEN(sBarcode) = 0 THEN
        _bRejected := TRUE;                                  // 空串拒入 / Empty barcode rejected
        _eCause := E_DL_EftCause.eBarcodeEmpty;              // 归因：条码空串（信息级） / Cause: empty barcode, info level
    ELSE
        (* 线性查重：扫描在队记录（带守护计数，深度有限故必然收敛） *)
        _bDup  := FALSE;                                     // 查重结论预置 / Duplicate result preset
        _uScan := 0;                                         // 扫描计数器归零 / Scan guard reset
        _iScanIdx := _iHead;                                 // 从当前头指针起扫 / Start at the current head
        WHILE (_uScan < DL_EFT_GUARD) AND (_uScan < _iCnt) DO
            IF aRec[_iScanIdx].sBarcode = sBarcode THEN
                _bDup := TRUE;                               // 命中重复条码 / Duplicate barcode found
            END_IF
            _uScan := _uScan + 1;                            // 计数器推进 / Guard advance
            _iScanIdx := _iScanIdx + 1;                      // 槽位推进 / Slot advance
            IF _iScanIdx > DL_EFT_DEPTH THEN
                _iScanIdx := 1;                              // 环形回卷 / Ring wrap
            END_IF
        END_WHILE

        IF _bDup THEN
            _bRejected := TRUE;                              // 重复条码拒入 / Duplicate barcode rejected
            _eCause := E_DL_EftCause.eDupBarcode;            // 归因：条码重复（信息级） / Cause: duplicate barcode, info level
        ELSIF _iCnt >= DL_EFT_DEPTH THEN
            _bRejected := TRUE;                              // 队满拒入 / Queue full, rejected
            _bFull := TRUE;                                  // 队满锁存（入队前判满语义） / Latch the full state
            _eCause := E_DL_EftCause.eQueueFull;             // 归因：队满 / Cause: queue full
        ELSE
            aRec[_iTail].sBatchNo  := sBatchNo;              // 写尾记录批次号 / Write the tail batch number
            aRec[_iTail].sBarcode  := sBarcode;              // 写尾记录条码 / Write the tail barcode
            aRec[_iTail].fVolumeMl := fVolumeMl;             // 写尾记录注液量 / Write the tail volume
            _iCnt  := _iCnt + 1;                             // 计数递增 / Count increment
            _iTail := _iTail + 1;                            // 尾指针推进 / Tail advance
            IF _iTail > DL_EFT_DEPTH THEN
                _iTail := 1;                                 // 环形回卷 / Ring wrap
            END_IF
        END_IF
    END_IF
END_IF

(* —— 段 7：出口单点映射（名实双出口，R191） —— *)
iQueueCnt   := _iCnt;                                        // 在队条数出口 / Queued count outlet
bOutValid   := _bOutValid;                                   // 出队脉冲出口 / Dequeue pulse outlet
bQueueFull  := _bFull;                                       // 队满出口 / Full outlet
bRejected   := _bRejected;                                   // 拒入标志出口 / Reject outlet
bFullRelease:= _bFullRel;                                    // 满解除脉冲出口 / Full-release outlet
eState      := _eState;                                      // 相出口 / Phase outlet
eCause      := _eCause;                                      // 成因出口 / Cause outlet
bError      := _bFault;                                      // 故障标志（仅故障级码置位） / Error flag, fault level only

END_FUNCTION_BLOCK
